(* IEC 61131-3 sources: Aqueous_Solutions/docs-authority/plc (part 2) *)

(* ---- PLC-FAB.st ---- *)
(* AQS-CTL-004 X-CTL-04: control program source, generated by flow_graph/control/plc_programs.py *)
(* Basis: AQS-CTL-001 INSTRUMENT_INDEX.csv, AQS-CTL-002 control architecture, graph set-points. *)
(* PLC-FAB: CPU single; IO counts AI 72 AO 3 DI 92 DO 13 (modules per AQS-CTL-002, 16-channel, 20 % spare) *)
PROGRAM PLC_FAB_CTRL
VAR
  (* 100 ms cyclic task per AQS-CTL-002 *)
  WAFER_FABFT-01_PV : REAL ;  (* S39 normal 0.14 L/h )
  WAFER_FABFT-02_PV : REAL ;  (* S39B normal 0.00 L/h )
  WAFER_FABFT-03_PV : REAL ;  (* IA-FAB-SPENT normal 2.77 L/h )
  WAFER_FABFT-04_PV : REAL ;  (* IA-FAB-N2-VENT normal 0.03 L/h )
  WAFER_FABFT-05_PV : REAL ;  (* IA-AR-CZ-BACK normal 0.14 L/h )
  WAFER_FABLT-01_PV : REAL ;  (* A-M-182 liquid height )
  WAFER_FABPT-01_PV : REAL ;  (* no design pressure on the graph )
  WAFER_FABTE-01_PV : REAL ;  (* band by service )
  WET_BENCHFT-01_PV : REAL ;  (* S10 normal 3.29 L/h )
  WET_BENCHFT-02_PV : REAL ;  (* S38 normal 0.00 L/h )
  WET_BENCHLT-01_PV : REAL ;  (* A-M-182 liquid height )
  WET_BENCHPT-01_PV : REAL ;  (* no design pressure on the graph )
  WET_BENCHTE-01_PV : REAL ;  (* band by service )
  LITHO_ALIGNPT-01_PV : REAL ;  (* no design pressure on the graph )
  LITHO_ALIGNTE-01_PV : REAL ;  (* band by service )
  LITHO_COATPT-01_PV : REAL ;  (* no design pressure on the graph )
  LITHO_COATTE-01_PV : REAL ;  (* band by service )
  RESIST_SYNLT-01_PV : REAL ;  (* A-M-182 liquid height )
  RESIST_SYNPT-01_PV : REAL ;  (* no design pressure on the graph )
  RESIST_SYNTE-01_PV : REAL ;  (* band by service )
  SOLV_PLANTLT-01_PV : REAL ;  (* A-M-182 liquid height )
  SOLV_PLANTPT-01_PV : REAL ;  (* no design pressure on the graph )
  SOLV_PLANTTE-01_PV : REAL ;  (* band by service )
  WS_AMMONIAFT-01_PV : REAL ;  (* S33 normal 0.13 L/h )
  WS_AMMONIAFT-02_PV : REAL ;  (* IA-NH3-MET normal 0.00 L/h )
  WS_AMMONIALT-01_PV : REAL ;  (* A-M-182 liquid height )
  WS_AMMONIAPT-01_PV : REAL ;  (* no design pressure on the graph )
  WS_AMMONIATE-01_PV : REAL ;  (* band by service )
  WS_DOPELT-01_PV : REAL ;  (* A-M-182 liquid height )
  WS_DOPEPT-01_PV : REAL ;  (* no design pressure on the graph )
  WS_DOPETE-01_PV : REAL ;  (* band by service )
  WS_HF_EDFT-01_PV : REAL ;  (* S31 normal 0.06 L/h )
  WS_HF_EDLT-01_PV : REAL ;  (* A-M-182 liquid height )
  WS_HF_EDPT-01_PV : REAL ;  (* no design pressure on the graph )
  WS_HF_EDTE-01_PV : REAL ;  (* band by service )
  WS_KOHFT-01_PV : REAL ;  (* S35 normal 0.01 L/h )
  WS_KOHLT-01_PV : REAL ;  (* A-M-182 liquid height )
  WS_KOHPT-01_PV : REAL ;  (* no design pressure on the graph )
  WS_KOHTE-01_PV : REAL ;  (* band by service )
  WS_NITRICFT-01_PV : REAL ;  (* S34 normal 0.05 L/h )
  WS_NITRICFT-02_PV : REAL ;  (* IA-NIT-VENT normal 0.00 L/h )
  WS_NITRICLT-01_PV : REAL ;  (* A-M-182 liquid height )
  WS_NITRICPT-01_PV : REAL ;  (* no design pressure on the graph )
  WS_NITRICTE-01_PV : REAL ;  (* band by service )
  WS_PEROXFT-01_PV : REAL ;  (* S32 normal 0.12 L/h )
  WS_PEROXLT-01_PV : REAL ;  (* A-M-182 liquid height )
  WS_PEROXPT-01_PV : REAL ;  (* no design pressure on the graph )
  WS_PEROXTE-01_PV : REAL ;  (* band by service )
  WS_PHOSFT-01_PV : REAL ;  (* S34B normal 0.03 L/h )
  WS_PHOSFT-02_PV : REAL ;  (* IA-PHOS-DOPE normal 0.00 L/h )
  WS_PHOSLT-01_PV : REAL ;  (* A-M-182 liquid height )
  WS_PHOSPT-01_PV : REAL ;  (* no design pressure on the graph )
  WS_PHOSTE-01_PV : REAL ;  (* band by service )
  WS_SLURRYFT-01_PV : REAL ;  (* S37 normal 0.14 L/h )
  WS_SLURRYLT-01_PV : REAL ;  (* A-M-182 liquid height )
  WS_SLURRYPT-01_PV : REAL ;  (* no design pressure on the graph )
  WS_SLURRYTE-01_PV : REAL ;  (* band by service )
  WS_SOLVFT-01_PV : REAL ;  (* IA-SOLV-WB normal 0.01 L/h )
  WS_SOLVFT-02_PV : REAL ;  (* IA-FAB-SOLV normal 0.00 L/h )
  WS_SOLVLT-01_PV : REAL ;  (* A-M-182 liquid height )
  WS_SOLVPT-01_PV : REAL ;  (* no design pressure on the graph )
  WS_SOLVTE-01_PV : REAL ;  (* band by service )
  LITHO_STUBPT-01_PV : REAL ;  (* no design pressure on the graph )
  LITHO_STUBTE-01_PV : REAL ;  (* band by service )
  FAB_UPW_TANKFT-01_PV : REAL ;  (* S27 normal 2.50 L/h )
  FAB_UPW_TANKLT-01_PV : REAL ;  (* A-M-182 liquid height )
  FAB_UPW_TANKPT-01_PV : REAL ;  (* no design pressure on the graph )
  FAB_UPW_TANKTE-01_PV : REAL ;  (* band by service )
  SOLAR_PV_CELLPT-01_PV : REAL ;  (* no design pressure on the graph )
  SOLAR_PV_CELLTE-01_PV : REAL ;  (* band by service )
  LITHO_DEVPT-01_PV : REAL ;  (* no design pressure on the graph )
  LITHO_DEVTE-01_PV : REAL ;  (* band by service )
END_VAR

  (* FLOW control loop - set-point from the graph basis *)
  WAFER_FABFT-01_SP := 0.14 ;  (* graph basis: S39 normal 0.14 L/h )
  FB_PI_WAFER_FABFT-01( PV := WAFER_FABFT-01_PV, SP := WAFER_FABFT-01_SP );  (* PI per AQS-CTL-002; GAIN/KI entered at commissioning from the step test (AQS-COM-001 sec. 3), anti-windup clamp per this FB *)
  WAFER_FABFT-01_ALARM_HI := 0.15400000000000003 ;  (* SP x 1.1 margin, A-M-188 margin class *)
  WAFER_FABFT-01_ALARM_LO := 0.12600000000000003 ;

  (* FLOW control loop - set-point from the graph basis *)
  WAFER_FABFT-02_SP := 0.0 ;  (* graph basis: S39B normal 0.00 L/h )
  FB_PI_WAFER_FABFT-02( PV := WAFER_FABFT-02_PV, SP := WAFER_FABFT-02_SP );  (* PI per AQS-CTL-002; GAIN/KI entered at commissioning from the step test (AQS-COM-001 sec. 3), anti-windup clamp per this FB *)
  WAFER_FABFT-02_ALARM_HI := 0.0 ;  (* expected-zero state: any positive PV alarms )

  (* FLOW control loop - set-point from the graph basis *)
  WAFER_FABFT-03_SP := 2.77 ;  (* graph basis: IA-FAB-SPENT normal 2.77 L/h )
  FB_PI_WAFER_FABFT-03( PV := WAFER_FABFT-03_PV, SP := WAFER_FABFT-03_SP );  (* PI per AQS-CTL-002; GAIN/KI entered at commissioning from the step test (AQS-COM-001 sec. 3), anti-windup clamp per this FB *)
  WAFER_FABFT-03_ALARM_HI := 3.047 ;  (* SP x 1.1 margin, A-M-188 margin class *)
  WAFER_FABFT-03_ALARM_LO := 2.493 ;

  (* FLOW control loop - set-point from the graph basis *)
  WAFER_FABFT-04_SP := 0.03 ;  (* graph basis: IA-FAB-N2-VENT normal 0.03 L/h )
  FB_PI_WAFER_FABFT-04( PV := WAFER_FABFT-04_PV, SP := WAFER_FABFT-04_SP );  (* PI per AQS-CTL-002; GAIN/KI entered at commissioning from the step test (AQS-COM-001 sec. 3), anti-windup clamp per this FB *)
  WAFER_FABFT-04_ALARM_HI := 0.033 ;  (* SP x 1.1 margin, A-M-188 margin class *)
  WAFER_FABFT-04_ALARM_LO := 0.027 ;

  (* FLOW control loop - set-point from the graph basis *)
  WAFER_FABFT-05_SP := 0.14 ;  (* graph basis: IA-AR-CZ-BACK normal 0.14 L/h )
  FB_PI_WAFER_FABFT-05( PV := WAFER_FABFT-05_PV, SP := WAFER_FABFT-05_SP );  (* PI per AQS-CTL-002; GAIN/KI entered at commissioning from the step test (AQS-COM-001 sec. 3), anti-windup clamp per this FB *)
  WAFER_FABFT-05_ALARM_HI := 0.15400000000000003 ;  (* SP x 1.1 margin, A-M-188 margin class *)
  WAFER_FABFT-05_ALARM_LO := 0.12600000000000003 ;

  (* LEVEL monitoring block - indication, no set-point invented )
  FB_AI_WAFER_FABLT-01( PV := WAFER_FABLT-01_PV );
  WAFER_FABLT-01_ALARM_HI := 90.0 ;  (* 90 % of span, registered LSH convention )

  (* PRESSURE monitoring block - indication, no set-point invented )
  FB_AI_WAFER_FABPT-01( PV := WAFER_FABPT-01_PV );
  WAFER_FABPT-01_ALARM_HI := 9.0 ;  (* 90 % of span, registered LSH convention )

  (* TEMPERATURE monitoring block - indication, no set-point invented )
  FB_AI_WAFER_FABTE-01( PV := WAFER_FABTE-01_PV );
  WAFER_FABTE-01_ALARM_HI := 135.0 ;  (* 90 % of span, registered LSH convention )

  (* FLOW control loop - set-point from the graph basis *)
  WET_BENCHFT-01_SP := 3.29 ;  (* graph basis: S10 normal 3.29 L/h )
  FB_PI_WET_BENCHFT-01( PV := WET_BENCHFT-01_PV, SP := WET_BENCHFT-01_SP );  (* PI per AQS-CTL-002; GAIN/KI entered at commissioning from the step test (AQS-COM-001 sec. 3), anti-windup clamp per this FB *)
  WET_BENCHFT-01_ALARM_HI := 3.619 ;  (* SP x 1.1 margin, A-M-188 margin class *)
  WET_BENCHFT-01_ALARM_LO := 2.9610000000000003 ;

  (* FLOW control loop - set-point from the graph basis *)
  WET_BENCHFT-02_SP := 0.0 ;  (* graph basis: S38 normal 0.00 L/h )
  FB_PI_WET_BENCHFT-02( PV := WET_BENCHFT-02_PV, SP := WET_BENCHFT-02_SP );  (* PI per AQS-CTL-002; GAIN/KI entered at commissioning from the step test (AQS-COM-001 sec. 3), anti-windup clamp per this FB *)
  WET_BENCHFT-02_ALARM_HI := 0.0 ;  (* expected-zero state: any positive PV alarms )

  (* LEVEL monitoring block - indication, no set-point invented )
  FB_AI_WET_BENCHLT-01( PV := WET_BENCHLT-01_PV );
  WET_BENCHLT-01_ALARM_HI := 90.0 ;  (* 90 % of span, registered LSH convention )

  (* PRESSURE monitoring block - indication, no set-point invented )
  FB_AI_WET_BENCHPT-01( PV := WET_BENCHPT-01_PV );
  WET_BENCHPT-01_ALARM_HI := 9.0 ;  (* 90 % of span, registered LSH convention )

  (* TEMPERATURE monitoring block - indication, no set-point invented )
  FB_AI_WET_BENCHTE-01( PV := WET_BENCHTE-01_PV );
  WET_BENCHTE-01_ALARM_HI := 135.0 ;  (* 90 % of span, registered LSH convention )

  (* PRESSURE monitoring block - indication, no set-point invented )
  FB_AI_LITHO_ALIGNPT-01( PV := LITHO_ALIGNPT-01_PV );
  LITHO_ALIGNPT-01_ALARM_HI := 9.0 ;  (* 90 % of span, registered LSH convention )

  (* TEMPERATURE monitoring block - indication, no set-point invented )
  FB_AI_LITHO_ALIGNTE-01( PV := LITHO_ALIGNTE-01_PV );
  LITHO_ALIGNTE-01_ALARM_HI := 135.0 ;  (* 90 % of span, registered LSH convention )

  (* PRESSURE monitoring block - indication, no set-point invented )
  FB_AI_LITHO_COATPT-01( PV := LITHO_COATPT-01_PV );
  LITHO_COATPT-01_ALARM_HI := 9.0 ;  (* 90 % of span, registered LSH convention )

  (* TEMPERATURE monitoring block - indication, no set-point invented )
  FB_AI_LITHO_COATTE-01( PV := LITHO_COATTE-01_PV );
  LITHO_COATTE-01_ALARM_HI := 135.0 ;  (* 90 % of span, registered LSH convention )

  (* LEVEL monitoring block - indication, no set-point invented )
  FB_AI_RESIST_SYNLT-01( PV := RESIST_SYNLT-01_PV );
  RESIST_SYNLT-01_ALARM_HI := 90.0 ;  (* 90 % of span, registered LSH convention )

  (* PRESSURE monitoring block - indication, no set-point invented )
  FB_AI_RESIST_SYNPT-01( PV := RESIST_SYNPT-01_PV );
  RESIST_SYNPT-01_ALARM_HI := 9.0 ;  (* 90 % of span, registered LSH convention )

  (* TEMPERATURE monitoring block - indication, no set-point invented )
  FB_AI_RESIST_SYNTE-01( PV := RESIST_SYNTE-01_PV );
  RESIST_SYNTE-01_ALARM_HI := 135.0 ;  (* 90 % of span, registered LSH convention )

  (* LEVEL monitoring block - indication, no set-point invented )
  FB_AI_SOLV_PLANTLT-01( PV := SOLV_PLANTLT-01_PV );
  SOLV_PLANTLT-01_ALARM_HI := 90.0 ;  (* 90 % of span, registered LSH convention )

  (* PRESSURE monitoring block - indication, no set-point invented )
  FB_AI_SOLV_PLANTPT-01( PV := SOLV_PLANTPT-01_PV );
  SOLV_PLANTPT-01_ALARM_HI := 9.0 ;  (* 90 % of span, registered LSH convention )

  (* TEMPERATURE monitoring block - indication, no set-point invented )
  FB_AI_SOLV_PLANTTE-01( PV := SOLV_PLANTTE-01_PV );
  SOLV_PLANTTE-01_ALARM_HI := 135.0 ;  (* 90 % of span, registered LSH convention )

  (* FLOW control loop - set-point from the graph basis *)
  WS_AMMONIAFT-01_SP := 0.13 ;  (* graph basis: S33 normal 0.13 L/h )
  FB_PI_WS_AMMONIAFT-01( PV := WS_AMMONIAFT-01_PV, SP := WS_AMMONIAFT-01_SP );  (* PI per AQS-CTL-002; GAIN/KI entered at commissioning from the step test (AQS-COM-001 sec. 3), anti-windup clamp per this FB *)
  WS_AMMONIAFT-01_ALARM_HI := 0.14300000000000002 ;  (* SP x 1.1 margin, A-M-188 margin class *)
  WS_AMMONIAFT-01_ALARM_LO := 0.117 ;

  (* FLOW control loop - set-point from the graph basis *)
  WS_AMMONIAFT-02_SP := 0.0 ;  (* graph basis: IA-NH3-MET normal 0.00 L/h )
  FB_PI_WS_AMMONIAFT-02( PV := WS_AMMONIAFT-02_PV, SP := WS_AMMONIAFT-02_SP );  (* PI per AQS-CTL-002; GAIN/KI entered at commissioning from the step test (AQS-COM-001 sec. 3), anti-windup clamp per this FB *)
  WS_AMMONIAFT-02_ALARM_HI := 0.0 ;  (* expected-zero state: any positive PV alarms )

  (* LEVEL monitoring block - indication, no set-point invented )
  FB_AI_WS_AMMONIALT-01( PV := WS_AMMONIALT-01_PV );
  WS_AMMONIALT-01_ALARM_HI := 90.0 ;  (* 90 % of span, registered LSH convention )

  (* PRESSURE monitoring block - indication, no set-point invented )
  FB_AI_WS_AMMONIAPT-01( PV := WS_AMMONIAPT-01_PV );
  WS_AMMONIAPT-01_ALARM_HI := 9.0 ;  (* 90 % of span, registered LSH convention )

  (* TEMPERATURE monitoring block - indication, no set-point invented )
  FB_AI_WS_AMMONIATE-01( PV := WS_AMMONIATE-01_PV );
  WS_AMMONIATE-01_ALARM_HI := 135.0 ;  (* 90 % of span, registered LSH convention )

  (* LEVEL monitoring block - indication, no set-point invented )
  FB_AI_WS_DOPELT-01( PV := WS_DOPELT-01_PV );
  WS_DOPELT-01_ALARM_HI := 90.0 ;  (* 90 % of span, registered LSH convention )

  (* PRESSURE monitoring block - indication, no set-point invented )
  FB_AI_WS_DOPEPT-01( PV := WS_DOPEPT-01_PV );
  WS_DOPEPT-01_ALARM_HI := 9.0 ;  (* 90 % of span, registered LSH convention )

  (* TEMPERATURE monitoring block - indication, no set-point invented )
  FB_AI_WS_DOPETE-01( PV := WS_DOPETE-01_PV );
  WS_DOPETE-01_ALARM_HI := 135.0 ;  (* 90 % of span, registered LSH convention )

  (* FLOW control loop - set-point from the graph basis *)
  WS_HF_EDFT-01_SP := 0.06 ;  (* graph basis: S31 normal 0.06 L/h )
  FB_PI_WS_HF_EDFT-01( PV := WS_HF_EDFT-01_PV, SP := WS_HF_EDFT-01_SP );  (* PI per AQS-CTL-002; GAIN/KI entered at commissioning from the step test (AQS-COM-001 sec. 3), anti-windup clamp per this FB *)
  WS_HF_EDFT-01_ALARM_HI := 0.066 ;  (* SP x 1.1 margin, A-M-188 margin class *)
  WS_HF_EDFT-01_ALARM_LO := 0.054 ;

  (* LEVEL monitoring block - indication, no set-point invented )
  FB_AI_WS_HF_EDLT-01( PV := WS_HF_EDLT-01_PV );
  WS_HF_EDLT-01_ALARM_HI := 90.0 ;  (* 90 % of span, registered LSH convention )

  (* PRESSURE monitoring block - indication, no set-point invented )
  FB_AI_WS_HF_EDPT-01( PV := WS_HF_EDPT-01_PV );
  WS_HF_EDPT-01_ALARM_HI := 9.0 ;  (* 90 % of span, registered LSH convention )

  (* TEMPERATURE monitoring block - indication, no set-point invented )
  FB_AI_WS_HF_EDTE-01( PV := WS_HF_EDTE-01_PV );
  WS_HF_EDTE-01_ALARM_HI := 135.0 ;  (* 90 % of span, registered LSH convention )

  (* FLOW control loop - set-point from the graph basis *)
  WS_KOHFT-01_SP := 0.01 ;  (* graph basis: S35 normal 0.01 L/h )
  FB_PI_WS_KOHFT-01( PV := WS_KOHFT-01_PV, SP := WS_KOHFT-01_SP );  (* PI per AQS-CTL-002; GAIN/KI entered at commissioning from the step test (AQS-COM-001 sec. 3), anti-windup clamp per this FB *)
  WS_KOHFT-01_ALARM_HI := 0.011000000000000001 ;  (* SP x 1.1 margin, A-M-188 margin class *)
  WS_KOHFT-01_ALARM_LO := 0.009000000000000001 ;

  (* LEVEL monitoring block - indication, no set-point invented )
  FB_AI_WS_KOHLT-01( PV := WS_KOHLT-01_PV );
  WS_KOHLT-01_ALARM_HI := 90.0 ;  (* 90 % of span, registered LSH convention )

  (* PRESSURE monitoring block - indication, no set-point invented )
  FB_AI_WS_KOHPT-01( PV := WS_KOHPT-01_PV );
  WS_KOHPT-01_ALARM_HI := 9.0 ;  (* 90 % of span, registered LSH convention )

  (* TEMPERATURE monitoring block - indication, no set-point invented )
  FB_AI_WS_KOHTE-01( PV := WS_KOHTE-01_PV );
  WS_KOHTE-01_ALARM_HI := 135.0 ;  (* 90 % of span, registered LSH convention )

  (* FLOW control loop - set-point from the graph basis *)
  WS_NITRICFT-01_SP := 0.05 ;  (* graph basis: S34 normal 0.05 L/h )
  FB_PI_WS_NITRICFT-01( PV := WS_NITRICFT-01_PV, SP := WS_NITRICFT-01_SP );  (* PI per AQS-CTL-002; GAIN/KI entered at commissioning from the step test (AQS-COM-001 sec. 3), anti-windup clamp per this FB *)
  WS_NITRICFT-01_ALARM_HI := 0.05500000000000001 ;  (* SP x 1.1 margin, A-M-188 margin class *)
  WS_NITRICFT-01_ALARM_LO := 0.045000000000000005 ;

  (* FLOW control loop - set-point from the graph basis *)
  WS_NITRICFT-02_SP := 0.0 ;  (* graph basis: IA-NIT-VENT normal 0.00 L/h )
  FB_PI_WS_NITRICFT-02( PV := WS_NITRICFT-02_PV, SP := WS_NITRICFT-02_SP );  (* PI per AQS-CTL-002; GAIN/KI entered at commissioning from the step test (AQS-COM-001 sec. 3), anti-windup clamp per this FB *)
  WS_NITRICFT-02_ALARM_HI := 0.0 ;  (* expected-zero state: any positive PV alarms )

  (* LEVEL monitoring block - indication, no set-point invented )
  FB_AI_WS_NITRICLT-01( PV := WS_NITRICLT-01_PV );
  WS_NITRICLT-01_ALARM_HI := 90.0 ;  (* 90 % of span, registered LSH convention )

  (* PRESSURE monitoring block - indication, no set-point invented )
  FB_AI_WS_NITRICPT-01( PV := WS_NITRICPT-01_PV );
  WS_NITRICPT-01_ALARM_HI := 9.0 ;  (* 90 % of span, registered LSH convention )

  (* TEMPERATURE monitoring block - indication, no set-point invented )
  FB_AI_WS_NITRICTE-01( PV := WS_NITRICTE-01_PV );
  WS_NITRICTE-01_ALARM_HI := 135.0 ;  (* 90 % of span, registered LSH convention )

  (* FLOW control loop - set-point from the graph basis *)
  WS_PEROXFT-01_SP := 0.12 ;  (* graph basis: S32 normal 0.12 L/h )
  FB_PI_WS_PEROXFT-01( PV := WS_PEROXFT-01_PV, SP := WS_PEROXFT-01_SP );  (* PI per AQS-CTL-002; GAIN/KI entered at commissioning from the step test (AQS-COM-001 sec. 3), anti-windup clamp per this FB *)
  WS_PEROXFT-01_ALARM_HI := 0.132 ;  (* SP x 1.1 margin, A-M-188 margin class *)
  WS_PEROXFT-01_ALARM_LO := 0.108 ;

  (* LEVEL monitoring block - indication, no set-point invented )
  FB_AI_WS_PEROXLT-01( PV := WS_PEROXLT-01_PV );
  WS_PEROXLT-01_ALARM_HI := 90.0 ;  (* 90 % of span, registered LSH convention )

  (* PRESSURE monitoring block - indication, no set-point invented )
  FB_AI_WS_PEROXPT-01( PV := WS_PEROXPT-01_PV );
  WS_PEROXPT-01_ALARM_HI := 9.0 ;  (* 90 % of span, registered LSH convention )

  (* TEMPERATURE monitoring block - indication, no set-point invented )
  FB_AI_WS_PEROXTE-01( PV := WS_PEROXTE-01_PV );
  WS_PEROXTE-01_ALARM_HI := 135.0 ;  (* 90 % of span, registered LSH convention )

  (* FLOW control loop - set-point from the graph basis *)
  WS_PHOSFT-01_SP := 0.03 ;  (* graph basis: S34B normal 0.03 L/h )
  FB_PI_WS_PHOSFT-01( PV := WS_PHOSFT-01_PV, SP := WS_PHOSFT-01_SP );  (* PI per AQS-CTL-002; GAIN/KI entered at commissioning from the step test (AQS-COM-001 sec. 3), anti-windup clamp per this FB *)
  WS_PHOSFT-01_ALARM_HI := 0.033 ;  (* SP x 1.1 margin, A-M-188 margin class *)
  WS_PHOSFT-01_ALARM_LO := 0.027 ;

  (* FLOW control loop - set-point from the graph basis *)
  WS_PHOSFT-02_SP := 0.0 ;  (* graph basis: IA-PHOS-DOPE normal 0.00 L/h )
  FB_PI_WS_PHOSFT-02( PV := WS_PHOSFT-02_PV, SP := WS_PHOSFT-02_SP );  (* PI per AQS-CTL-002; GAIN/KI entered at commissioning from the step test (AQS-COM-001 sec. 3), anti-windup clamp per this FB *)
  WS_PHOSFT-02_ALARM_HI := 0.0 ;  (* expected-zero state: any positive PV alarms )

  (* LEVEL monitoring block - indication, no set-point invented )
  FB_AI_WS_PHOSLT-01( PV := WS_PHOSLT-01_PV );
  WS_PHOSLT-01_ALARM_HI := 90.0 ;  (* 90 % of span, registered LSH convention )

  (* PRESSURE monitoring block - indication, no set-point invented )
  FB_AI_WS_PHOSPT-01( PV := WS_PHOSPT-01_PV );
  WS_PHOSPT-01_ALARM_HI := 9.0 ;  (* 90 % of span, registered LSH convention )

  (* TEMPERATURE monitoring block - indication, no set-point invented )
  FB_AI_WS_PHOSTE-01( PV := WS_PHOSTE-01_PV );
  WS_PHOSTE-01_ALARM_HI := 135.0 ;  (* 90 % of span, registered LSH convention )

  (* FLOW control loop - set-point from the graph basis *)
  WS_SLURRYFT-01_SP := 0.14 ;  (* graph basis: S37 normal 0.14 L/h )
  FB_PI_WS_SLURRYFT-01( PV := WS_SLURRYFT-01_PV, SP := WS_SLURRYFT-01_SP );  (* PI per AQS-CTL-002; GAIN/KI entered at commissioning from the step test (AQS-COM-001 sec. 3), anti-windup clamp per this FB *)
  WS_SLURRYFT-01_ALARM_HI := 0.15400000000000003 ;  (* SP x 1.1 margin, A-M-188 margin class *)
  WS_SLURRYFT-01_ALARM_LO := 0.12600000000000003 ;

  (* LEVEL monitoring block - indication, no set-point invented )
  FB_AI_WS_SLURRYLT-01( PV := WS_SLURRYLT-01_PV );
  WS_SLURRYLT-01_ALARM_HI := 90.0 ;  (* 90 % of span, registered LSH convention )

  (* PRESSURE monitoring block - indication, no set-point invented )
  FB_AI_WS_SLURRYPT-01( PV := WS_SLURRYPT-01_PV );
  WS_SLURRYPT-01_ALARM_HI := 9.0 ;  (* 90 % of span, registered LSH convention )

  (* TEMPERATURE monitoring block - indication, no set-point invented )
  FB_AI_WS_SLURRYTE-01( PV := WS_SLURRYTE-01_PV );
  WS_SLURRYTE-01_ALARM_HI := 135.0 ;  (* 90 % of span, registered LSH convention )

  (* FLOW control loop - set-point from the graph basis *)
  WS_SOLVFT-01_SP := 0.01 ;  (* graph basis: IA-SOLV-WB normal 0.01 L/h )
  FB_PI_WS_SOLVFT-01( PV := WS_SOLVFT-01_PV, SP := WS_SOLVFT-01_SP );  (* PI per AQS-CTL-002; GAIN/KI entered at commissioning from the step test (AQS-COM-001 sec. 3), anti-windup clamp per this FB *)
  WS_SOLVFT-01_ALARM_HI := 0.011000000000000001 ;  (* SP x 1.1 margin, A-M-188 margin class *)
  WS_SOLVFT-01_ALARM_LO := 0.009000000000000001 ;

  (* FLOW control loop - set-point from the graph basis *)
  WS_SOLVFT-02_SP := 0.0 ;  (* graph basis: IA-FAB-SOLV normal 0.00 L/h )
  FB_PI_WS_SOLVFT-02( PV := WS_SOLVFT-02_PV, SP := WS_SOLVFT-02_SP );  (* PI per AQS-CTL-002; GAIN/KI entered at commissioning from the step test (AQS-COM-001 sec. 3), anti-windup clamp per this FB *)
  WS_SOLVFT-02_ALARM_HI := 0.0 ;  (* expected-zero state: any positive PV alarms )

  (* LEVEL monitoring block - indication, no set-point invented )
  FB_AI_WS_SOLVLT-01( PV := WS_SOLVLT-01_PV );
  WS_SOLVLT-01_ALARM_HI := 90.0 ;  (* 90 % of span, registered LSH convention )

  (* PRESSURE monitoring block - indication, no set-point invented )
  FB_AI_WS_SOLVPT-01( PV := WS_SOLVPT-01_PV );
  WS_SOLVPT-01_ALARM_HI := 9.0 ;  (* 90 % of span, registered LSH convention )

  (* TEMPERATURE monitoring block - indication, no set-point invented )
  FB_AI_WS_SOLVTE-01( PV := WS_SOLVTE-01_PV );
  WS_SOLVTE-01_ALARM_HI := 135.0 ;  (* 90 % of span, registered LSH convention )

  (* PRESSURE monitoring block - indication, no set-point invented )
  FB_AI_LITHO_STUBPT-01( PV := LITHO_STUBPT-01_PV );
  LITHO_STUBPT-01_ALARM_HI := 9.0 ;  (* 90 % of span, registered LSH convention )

  (* TEMPERATURE monitoring block - indication, no set-point invented )
  FB_AI_LITHO_STUBTE-01( PV := LITHO_STUBTE-01_PV );
  LITHO_STUBTE-01_ALARM_HI := 135.0 ;  (* 90 % of span, registered LSH convention )

  (* FLOW control loop - set-point from the graph basis *)
  FAB_UPW_TANKFT-01_SP := 2.5 ;  (* graph basis: S27 normal 2.50 L/h )
  FB_PI_FAB_UPW_TANKFT-01( PV := FAB_UPW_TANKFT-01_PV, SP := FAB_UPW_TANKFT-01_SP );  (* PI per AQS-CTL-002; GAIN/KI entered at commissioning from the step test (AQS-COM-001 sec. 3), anti-windup clamp per this FB *)
  FAB_UPW_TANKFT-01_ALARM_HI := 2.75 ;  (* SP x 1.1 margin, A-M-188 margin class *)
  FAB_UPW_TANKFT-01_ALARM_LO := 2.25 ;

  (* LEVEL monitoring block - indication, no set-point invented )
  FB_AI_FAB_UPW_TANKLT-01( PV := FAB_UPW_TANKLT-01_PV );
  FAB_UPW_TANKLT-01_ALARM_HI := 90.0 ;  (* 90 % of span, registered LSH convention )

  (* PRESSURE monitoring block - indication, no set-point invented )
  FB_AI_FAB_UPW_TANKPT-01( PV := FAB_UPW_TANKPT-01_PV );
  FAB_UPW_TANKPT-01_ALARM_HI := 9.0 ;  (* 90 % of span, registered LSH convention )

  (* TEMPERATURE monitoring block - indication, no set-point invented )
  FB_AI_FAB_UPW_TANKTE-01( PV := FAB_UPW_TANKTE-01_PV );
  FAB_UPW_TANKTE-01_ALARM_HI := 135.0 ;  (* 90 % of span, registered LSH convention )

  (* PRESSURE monitoring block - indication, no set-point invented )
  FB_AI_SOLAR_PV_CELLPT-01( PV := SOLAR_PV_CELLPT-01_PV );
  SOLAR_PV_CELLPT-01_ALARM_HI := 9.0 ;  (* 90 % of span, registered LSH convention )

  (* TEMPERATURE monitoring block - indication, no set-point invented )
  FB_AI_SOLAR_PV_CELLTE-01( PV := SOLAR_PV_CELLTE-01_PV );
  SOLAR_PV_CELLTE-01_ALARM_HI := 135.0 ;  (* 90 % of span, registered LSH convention )

  (* PRESSURE monitoring block - indication, no set-point invented )
  FB_AI_LITHO_DEVPT-01( PV := LITHO_DEVPT-01_PV );
  LITHO_DEVPT-01_ALARM_HI := 9.0 ;  (* 90 % of span, registered LSH convention )

  (* TEMPERATURE monitoring block - indication, no set-point invented )
  FB_AI_LITHO_DEVTE-01( PV := LITHO_DEVTE-01_PV );
  LITHO_DEVTE-01_ALARM_HI := 135.0 ;  (* 90 % of span, registered LSH convention )

END_PROGRAM

(* ---- PLC-FARM.st ---- *)
(* AQS-CTL-004 X-CTL-04: control program source, generated by flow_graph/control/plc_programs.py *)
(* Basis: AQS-CTL-001 INSTRUMENT_INDEX.csv, AQS-CTL-002 control architecture, graph set-points. *)
(* PLC-FARM: CPU redundant pair; IO counts AI 48 AO 0 DI 3 DO 0 (modules per AQS-CTL-002, 16-channel, 20 % spare) *)
PROGRAM PLC_FARM_CTRL
VAR
  (* 100 ms cyclic task per AQS-CTL-002 *)
  GROW_BEDFT-01_PV : REAL ;  (* S13 normal 0.16 L/h )
  GROW_BEDFT-02_PV : REAL ;  (* S15 normal 0.00 L/h )
  GROW_BEDFT-03_PV : REAL ;  (* S87 normal 0.03 L/h )
  GROW_BEDFT-04_PV : REAL ;  (* FARM_O2_TO_HAB normal 0.00 L/h )
  GROW_BEDFT-05_PV : REAL ;  (* IA-BED-VAP normal 2.81 L/h )
  GROW_BEDFT-06_PV : REAL ;  (* RABBIT_FORAGE normal 0.02 L/h )
  GROW_BEDFT-07_PV : REAL ;  (* NECTAR_FORAGE normal 0.01 L/h )
  GROW_BEDFT-08_PV : REAL ;  (* VERMI_FEED normal 0.04 L/h )
  GROW_BEDLT-01_PV : REAL ;  (* A-M-182 liquid height )
  GROW_BEDPT-01_PV : REAL ;  (* no design pressure on the graph )
  GROW_BEDTE-01_PV : REAL ;  (* band by service )
  DUCKWEEDPT-01_PV : REAL ;  (* no design pressure on the graph )
  DUCKWEEDTE-01_PV : REAL ;  (* band by service )
  BIOFILTERPT-01_PV : REAL ;  (* no design pressure on the graph )
  BIOFILTERTE-01_PV : REAL ;  (* band by service )
  BSFL_BINPT-01_PV : REAL ;  (* no design pressure on the graph )
  BSFL_BINTE-01_PV : REAL ;  (* band by service )
  QUAIL_CAGEPT-01_PV : REAL ;  (* no design pressure on the graph )
  QUAIL_CAGETE-01_PV : REAL ;  (* band by service )
  CHICKEN_COOPPT-01_PV : REAL ;  (* no design pressure on the graph )
  CHICKEN_COOPTE-01_PV : REAL ;  (* band by service )
  FEED_PREPPT-01_PV : REAL ;  (* no design pressure on the graph )
  FEED_PREPTE-01_PV : REAL ;  (* band by service )
  AQUA_TANKPT-01_PV : REAL ;  (* no design pressure on the graph )
  AQUA_TANKTE-01_PV : REAL ;  (* band by service )
  GROWBED_APT-01_PV : REAL ;  (* no design pressure on the graph )
  GROWBED_ATE-01_PV : REAL ;  (* band by service )
  GROWBED_BPT-01_PV : REAL ;  (* no design pressure on the graph )
  GROWBED_BTE-01_PV : REAL ;  (* band by service )
  BEE_HIVEPT-01_PV : REAL ;  (* no design pressure on the graph )
  BEE_HIVETE-01_PV : REAL ;  (* band by service )
  RABBIT_HUTCHPT-01_PV : REAL ;  (* no design pressure on the graph )
  RABBIT_HUTCHTE-01_PV : REAL ;  (* band by service )
  DUCK_PENPT-01_PV : REAL ;  (* no design pressure on the graph )
  DUCK_PENTE-01_PV : REAL ;  (* band by service )
  FOOD_STOREPT-01_PV : REAL ;  (* no design pressure on the graph )
  FOOD_STORETE-01_PV : REAL ;  (* band by service )
  AQUA_UVPT-01_PV : REAL ;  (* no design pressure on the graph )
  AQUA_UVTE-01_PV : REAL ;  (* band by service )
  VERMI_BINPT-01_PV : REAL ;  (* no design pressure on the graph )
  VERMI_BINTE-01_PV : REAL ;  (* band by service )
  FOOD_STORELT-01_PV : REAL ;  (* food stock level: S14 4.2 kg/d )
  HYDRO_GROWAE-01_PV : REAL ;  (* chamber CO2 watch against the habitat management set-point (X-LOC-10 placeholder )
  FEED_PREPPSH-01_PV : REAL ;  (* press-line overpressure interlock on the mash loop (X-FARM-10; A-M-426) )
  AQUA_UVFIT-01_PV : REAL ;  (* loop flow permissive: the UV dose is valid only above the minimum flow (X-FARM-1 )
  AQUA_UVUVT-01_PV : REAL ;  (* dose watchdog: lamp depletion or sleeve fouling decays the signal (X-FARM-12; A- )
  GROWBED_ALT-01_PV : REAL ;  (* flood-and-drain cycle watch on the aerobic root zone (X-FARM build-out; A-M-229) )
  GROWBED_BLT-01_PV : REAL ;  (* mineralisation-zone level watch (X-FARM build-out; A-M-229) )
END_VAR

  (* FLOW control loop - set-point from the graph basis *)
  GROW_BEDFT-01_SP := 0.16 ;  (* graph basis: S13 normal 0.16 L/h )
  FB_PI_GROW_BEDFT-01( PV := GROW_BEDFT-01_PV, SP := GROW_BEDFT-01_SP );  (* PI per AQS-CTL-002; GAIN/KI entered at commissioning from the step test (AQS-COM-001 sec. 3), anti-windup clamp per this FB *)
  GROW_BEDFT-01_ALARM_HI := 0.17600000000000002 ;  (* SP x 1.1 margin, A-M-188 margin class *)
  GROW_BEDFT-01_ALARM_LO := 0.14400000000000002 ;

  (* FLOW control loop - set-point from the graph basis *)
  GROW_BEDFT-02_SP := 0.0 ;  (* graph basis: S15 normal 0.00 L/h )
  FB_PI_GROW_BEDFT-02( PV := GROW_BEDFT-02_PV, SP := GROW_BEDFT-02_SP );  (* PI per AQS-CTL-002; GAIN/KI entered at commissioning from the step test (AQS-COM-001 sec. 3), anti-windup clamp per this FB *)
  GROW_BEDFT-02_ALARM_HI := 0.0 ;  (* expected-zero state: any positive PV alarms )

  (* FLOW control loop - set-point from the graph basis *)
  GROW_BEDFT-03_SP := 0.03 ;  (* graph basis: S87 normal 0.03 L/h )
  FB_PI_GROW_BEDFT-03( PV := GROW_BEDFT-03_PV, SP := GROW_BEDFT-03_SP );  (* PI per AQS-CTL-002; GAIN/KI entered at commissioning from the step test (AQS-COM-001 sec. 3), anti-windup clamp per this FB *)
  GROW_BEDFT-03_ALARM_HI := 0.033 ;  (* SP x 1.1 margin, A-M-188 margin class *)
  GROW_BEDFT-03_ALARM_LO := 0.027 ;

  (* FLOW control loop - set-point from the graph basis *)
  GROW_BEDFT-04_SP := 0.0 ;  (* graph basis: FARM_O2_TO_HAB normal 0.00 L/h )
  FB_PI_GROW_BEDFT-04( PV := GROW_BEDFT-04_PV, SP := GROW_BEDFT-04_SP );  (* PI per AQS-CTL-002; GAIN/KI entered at commissioning from the step test (AQS-COM-001 sec. 3), anti-windup clamp per this FB *)
  GROW_BEDFT-04_ALARM_HI := 0.0 ;  (* expected-zero state: any positive PV alarms )

  (* FLOW control loop - set-point from the graph basis *)
  GROW_BEDFT-05_SP := 2.81 ;  (* graph basis: IA-BED-VAP normal 2.81 L/h )
  FB_PI_GROW_BEDFT-05( PV := GROW_BEDFT-05_PV, SP := GROW_BEDFT-05_SP );  (* PI per AQS-CTL-002; GAIN/KI entered at commissioning from the step test (AQS-COM-001 sec. 3), anti-windup clamp per this FB *)
  GROW_BEDFT-05_ALARM_HI := 3.091 ;  (* SP x 1.1 margin, A-M-188 margin class *)
  GROW_BEDFT-05_ALARM_LO := 2.529 ;

  (* FLOW control loop - set-point from the graph basis *)
  GROW_BEDFT-06_SP := 0.02 ;  (* graph basis: RABBIT_FORAGE normal 0.02 L/h )
  FB_PI_GROW_BEDFT-06( PV := GROW_BEDFT-06_PV, SP := GROW_BEDFT-06_SP );  (* PI per AQS-CTL-002; GAIN/KI entered at commissioning from the step test (AQS-COM-001 sec. 3), anti-windup clamp per this FB *)
  GROW_BEDFT-06_ALARM_HI := 0.022000000000000002 ;  (* SP x 1.1 margin, A-M-188 margin class *)
  GROW_BEDFT-06_ALARM_LO := 0.018000000000000002 ;

  (* FLOW control loop - set-point from the graph basis *)
  GROW_BEDFT-07_SP := 0.01 ;  (* graph basis: NECTAR_FORAGE normal 0.01 L/h )
  FB_PI_GROW_BEDFT-07( PV := GROW_BEDFT-07_PV, SP := GROW_BEDFT-07_SP );  (* PI per AQS-CTL-002; GAIN/KI entered at commissioning from the step test (AQS-COM-001 sec. 3), anti-windup clamp per this FB *)
  GROW_BEDFT-07_ALARM_HI := 0.011000000000000001 ;  (* SP x 1.1 margin, A-M-188 margin class *)
  GROW_BEDFT-07_ALARM_LO := 0.009000000000000001 ;

  (* FLOW control loop - set-point from the graph basis *)
  GROW_BEDFT-08_SP := 0.04 ;  (* graph basis: VERMI_FEED normal 0.04 L/h )
  FB_PI_GROW_BEDFT-08( PV := GROW_BEDFT-08_PV, SP := GROW_BEDFT-08_SP );  (* PI per AQS-CTL-002; GAIN/KI entered at commissioning from the step test (AQS-COM-001 sec. 3), anti-windup clamp per this FB *)
  GROW_BEDFT-08_ALARM_HI := 0.044000000000000004 ;  (* SP x 1.1 margin, A-M-188 margin class *)
  GROW_BEDFT-08_ALARM_LO := 0.036000000000000004 ;

  (* LEVEL monitoring block - indication, no set-point invented )
  FB_AI_GROW_BEDLT-01( PV := GROW_BEDLT-01_PV );
  GROW_BEDLT-01_ALARM_HI := 90.0 ;  (* 90 % of span, registered LSH convention )

  (* PRESSURE monitoring block - indication, no set-point invented )
  FB_AI_GROW_BEDPT-01( PV := GROW_BEDPT-01_PV );
  GROW_BEDPT-01_ALARM_HI := 9.0 ;  (* 90 % of span, registered LSH convention )

  (* TEMPERATURE monitoring block - indication, no set-point invented )
  FB_AI_GROW_BEDTE-01( PV := GROW_BEDTE-01_PV );
  GROW_BEDTE-01_ALARM_HI := 135.0 ;  (* 90 % of span, registered LSH convention )

  (* PRESSURE monitoring block - indication, no set-point invented )
  FB_AI_DUCKWEEDPT-01( PV := DUCKWEEDPT-01_PV );
  DUCKWEEDPT-01_ALARM_HI := 9.0 ;  (* 90 % of span, registered LSH convention )

  (* TEMPERATURE monitoring block - indication, no set-point invented )
  FB_AI_DUCKWEEDTE-01( PV := DUCKWEEDTE-01_PV );
  DUCKWEEDTE-01_ALARM_HI := 135.0 ;  (* 90 % of span, registered LSH convention )

  (* PRESSURE monitoring block - indication, no set-point invented )
  FB_AI_BIOFILTERPT-01( PV := BIOFILTERPT-01_PV );
  BIOFILTERPT-01_ALARM_HI := 9.0 ;  (* 90 % of span, registered LSH convention )

  (* TEMPERATURE monitoring block - indication, no set-point invented )
  FB_AI_BIOFILTERTE-01( PV := BIOFILTERTE-01_PV );
  BIOFILTERTE-01_ALARM_HI := 135.0 ;  (* 90 % of span, registered LSH convention )

  (* PRESSURE monitoring block - indication, no set-point invented )
  FB_AI_BSFL_BINPT-01( PV := BSFL_BINPT-01_PV );
  BSFL_BINPT-01_ALARM_HI := 9.0 ;  (* 90 % of span, registered LSH convention )

  (* TEMPERATURE monitoring block - indication, no set-point invented )
  FB_AI_BSFL_BINTE-01( PV := BSFL_BINTE-01_PV );
  BSFL_BINTE-01_ALARM_HI := 135.0 ;  (* 90 % of span, registered LSH convention )

  (* PRESSURE monitoring block - indication, no set-point invented )
  FB_AI_QUAIL_CAGEPT-01( PV := QUAIL_CAGEPT-01_PV );
  QUAIL_CAGEPT-01_ALARM_HI := 9.0 ;  (* 90 % of span, registered LSH convention )

  (* TEMPERATURE monitoring block - indication, no set-point invented )
  FB_AI_QUAIL_CAGETE-01( PV := QUAIL_CAGETE-01_PV );
  QUAIL_CAGETE-01_ALARM_HI := 135.0 ;  (* 90 % of span, registered LSH convention )

  (* PRESSURE monitoring block - indication, no set-point invented )
  FB_AI_CHICKEN_COOPPT-01( PV := CHICKEN_COOPPT-01_PV );
  CHICKEN_COOPPT-01_ALARM_HI := 9.0 ;  (* 90 % of span, registered LSH convention )

  (* TEMPERATURE monitoring block - indication, no set-point invented )
  FB_AI_CHICKEN_COOPTE-01( PV := CHICKEN_COOPTE-01_PV );
  CHICKEN_COOPTE-01_ALARM_HI := 135.0 ;  (* 90 % of span, registered LSH convention )

  (* PRESSURE monitoring block - indication, no set-point invented )
  FB_AI_FEED_PREPPT-01( PV := FEED_PREPPT-01_PV );
  FEED_PREPPT-01_ALARM_HI := 9.0 ;  (* 90 % of span, registered LSH convention )

  (* TEMPERATURE monitoring block - indication, no set-point invented )
  FB_AI_FEED_PREPTE-01( PV := FEED_PREPTE-01_PV );
  FEED_PREPTE-01_ALARM_HI := 135.0 ;  (* 90 % of span, registered LSH convention )

  (* PRESSURE monitoring block - indication, no set-point invented )
  FB_AI_AQUA_TANKPT-01( PV := AQUA_TANKPT-01_PV );
  AQUA_TANKPT-01_ALARM_HI := 9.0 ;  (* 90 % of span, registered LSH convention )

  (* TEMPERATURE monitoring block - indication, no set-point invented )
  FB_AI_AQUA_TANKTE-01( PV := AQUA_TANKTE-01_PV );
  AQUA_TANKTE-01_ALARM_HI := 135.0 ;  (* 90 % of span, registered LSH convention )

  (* PRESSURE monitoring block - indication, no set-point invented )
  FB_AI_GROWBED_APT-01( PV := GROWBED_APT-01_PV );
  GROWBED_APT-01_ALARM_HI := 9.0 ;  (* 90 % of span, registered LSH convention )

  (* TEMPERATURE monitoring block - indication, no set-point invented )
  FB_AI_GROWBED_ATE-01( PV := GROWBED_ATE-01_PV );
  GROWBED_ATE-01_ALARM_HI := 135.0 ;  (* 90 % of span, registered LSH convention )

  (* PRESSURE monitoring block - indication, no set-point invented )
  FB_AI_GROWBED_BPT-01( PV := GROWBED_BPT-01_PV );
  GROWBED_BPT-01_ALARM_HI := 9.0 ;  (* 90 % of span, registered LSH convention )

  (* TEMPERATURE monitoring block - indication, no set-point invented )
  FB_AI_GROWBED_BTE-01( PV := GROWBED_BTE-01_PV );
  GROWBED_BTE-01_ALARM_HI := 135.0 ;  (* 90 % of span, registered LSH convention )

  (* PRESSURE monitoring block - indication, no set-point invented )
  FB_AI_BEE_HIVEPT-01( PV := BEE_HIVEPT-01_PV );
  BEE_HIVEPT-01_ALARM_HI := 9.0 ;  (* 90 % of span, registered LSH convention )

  (* TEMPERATURE monitoring block - indication, no set-point invented )
  FB_AI_BEE_HIVETE-01( PV := BEE_HIVETE-01_PV );
  BEE_HIVETE-01_ALARM_HI := 135.0 ;  (* 90 % of span, registered LSH convention )

  (* PRESSURE monitoring block - indication, no set-point invented )
  FB_AI_RABBIT_HUTCHPT-01( PV := RABBIT_HUTCHPT-01_PV );
  RABBIT_HUTCHPT-01_ALARM_HI := 9.0 ;  (* 90 % of span, registered LSH convention )

  (* TEMPERATURE monitoring block - indication, no set-point invented )
  FB_AI_RABBIT_HUTCHTE-01( PV := RABBIT_HUTCHTE-01_PV );
  RABBIT_HUTCHTE-01_ALARM_HI := 135.0 ;  (* 90 % of span, registered LSH convention )

  (* PRESSURE monitoring block - indication, no set-point invented )
  FB_AI_DUCK_PENPT-01( PV := DUCK_PENPT-01_PV );
  DUCK_PENPT-01_ALARM_HI := 9.0 ;  (* 90 % of span, registered LSH convention )

  (* TEMPERATURE monitoring block - indication, no set-point invented )
  FB_AI_DUCK_PENTE-01( PV := DUCK_PENTE-01_PV );
  DUCK_PENTE-01_ALARM_HI := 135.0 ;  (* 90 % of span, registered LSH convention )

  (* PRESSURE monitoring block - indication, no set-point invented )
  FB_AI_FOOD_STOREPT-01( PV := FOOD_STOREPT-01_PV );
  FOOD_STOREPT-01_ALARM_HI := 9.0 ;  (* 90 % of span, registered LSH convention )

  (* TEMPERATURE monitoring block - indication, no set-point invented )
  FB_AI_FOOD_STORETE-01( PV := FOOD_STORETE-01_PV );
  FOOD_STORETE-01_ALARM_HI := 135.0 ;  (* 90 % of span, registered LSH convention )

  (* PRESSURE monitoring block - indication, no set-point invented )
  FB_AI_AQUA_UVPT-01( PV := AQUA_UVPT-01_PV );
  AQUA_UVPT-01_ALARM_HI := 9.0 ;  (* 90 % of span, registered LSH convention )

  (* TEMPERATURE monitoring block - indication, no set-point invented )
  FB_AI_AQUA_UVTE-01( PV := AQUA_UVTE-01_PV );
  AQUA_UVTE-01_ALARM_HI := 135.0 ;  (* 90 % of span, registered LSH convention )

  (* PRESSURE monitoring block - indication, no set-point invented )
  FB_AI_VERMI_BINPT-01( PV := VERMI_BINPT-01_PV );
  VERMI_BINPT-01_ALARM_HI := 9.0 ;  (* 90 % of span, registered LSH convention )

  (* TEMPERATURE monitoring block - indication, no set-point invented )
  FB_AI_VERMI_BINTE-01( PV := VERMI_BINTE-01_PV );
  VERMI_BINTE-01_ALARM_HI := 135.0 ;  (* 90 % of span, registered LSH convention )

  (* LEVEL monitoring block - indication, no set-point invented )
  FB_AI_FOOD_STORELT-01( PV := FOOD_STORELT-01_PV );
  FOOD_STORELT-01_ALARM_HI := 90.0 ;  (* 90 % of span, registered LSH convention )

  (* CARBON-DIOXIDE monitoring block - indication, no set-point invented )
  FB_AI_HYDRO_GROWAE-01( PV := HYDRO_GROWAE-01_PV );
  HYDRO_GROWAE-01_ALARM_HI := 4500.0 ;  (* 90 % of span, registered LSH convention )

  (* PRESSURE monitoring block - indication, no set-point invented )
  FB_AI_FEED_PREPPSH-01( PV := FEED_PREPPSH-01_PV );
  FEED_PREPPSH-01_ALARM_HI := 225.0 ;  (* 90 % of span, registered LSH convention )

  (* FLOW monitoring block - indication, no set-point invented )
  FB_AI_AQUA_UVFIT-01( PV := AQUA_UVFIT-01_PV );
  AQUA_UVFIT-01_ALARM_HI := 90.0 ;  (* 90 % of span, registered LSH convention )

  (* UV monitoring block - indication, no set-point invented )
  FB_AI_AQUA_UVUVT-01( PV := AQUA_UVUVT-01_PV );
  AQUA_UVUVT-01_ALARM_HI := 4.5 ;  (* 90 % of span, registered LSH convention )

  (* LEVEL monitoring block - indication, no set-point invented )
  FB_AI_GROWBED_ALT-01( PV := GROWBED_ALT-01_PV );
  GROWBED_ALT-01_ALARM_HI := 270.0 ;  (* 90 % of span, registered LSH convention )

  (* LEVEL monitoring block - indication, no set-point invented )
  FB_AI_GROWBED_BLT-01( PV := GROWBED_BLT-01_PV );
  GROWBED_BLT-01_ALARM_HI := 270.0 ;  (* 90 % of span, registered LSH convention )

END_PROGRAM

(* ---- PLC-FOUNDRY.st ---- *)
(* AQS-CTL-004 X-CTL-04: control program source, generated by flow_graph/control/plc_programs.py *)
(* Basis: AQS-CTL-001 INSTRUMENT_INDEX.csv, AQS-CTL-002 control architecture, graph set-points. *)
(* PLC-FOUNDRY: CPU single; IO counts AI 87 AO 0 DI 19 DO 1 (modules per AQS-CTL-002, 16-channel, 20 % spare) *)
PROGRAM PLC_FOUNDRY_CTRL
VAR
  (* 100 ms cyclic task per AQS-CTL-002 *)
  AL_POTPT-01_PV : REAL ;  (* no design pressure on the graph )
  AL_POTTE-01_PV : REAL ;  (* band by service )
  CAST_LINELT-01_PV : REAL ;  (* A-M-182 liquid height )
  CAST_LINEPT-01_PV : REAL ;  (* no design pressure on the graph )
  CAST_LINETE-01_PV : REAL ;  (* band by service )
  CA_POTLT-01_PV : REAL ;  (* A-M-182 liquid height )
  CA_POTPT-01_PV : REAL ;  (* no design pressure on the graph )
  CA_POTTE-01_PV : REAL ;  (* band by service )
  COMB_HEATPT-01_PV : REAL ;  (* no design pressure on the graph )
  COMB_HEATTE-01_PV : REAL ;  (* band by service )
  CONT_CASTLT-01_PV : REAL ;  (* A-M-182 liquid height )
  CONT_CASTPT-01_PV : REAL ;  (* no design pressure on the graph )
  CONT_CASTTE-01_PV : REAL ;  (* band by service )
  CR_CELLPT-01_PV : REAL ;  (* no design pressure on the graph )
  CR_CELLTE-01_PV : REAL ;  (* band by service )
  DRAWPT-01_PV : REAL ;  (* no design pressure on the graph )
  DRAWTE-01_PV : REAL ;  (* band by service )
  EXTRUDEPT-01_PV : REAL ;  (* no design pressure on the graph )
  EXTRUDETE-01_PV : REAL ;  (* band by service )
  FLUX_PREPPT-01_PV : REAL ;  (* no design pressure on the graph )
  FLUX_PREPTE-01_PV : REAL ;  (* band by service )
  IND_MELTFT-01_PV : REAL ;  (* IND_MELT_TO_CAST normal 0.12 L/h )
  IND_MELTFT-02_PV : REAL ;  (* IND_TO_CONT normal 0.96 L/h )
  IND_MELTFT-03_PV : REAL ;  (* IND_TO_ATOM normal 0.00 L/h )
  IND_MELTFT-04_PV : REAL ;  (* IND_TO_INV normal 0.08 L/h )
  IND_MELTPT-01_PV : REAL ;  (* no design pressure on the graph )
  IND_MELTTE-01_PV : REAL ;  (* band by service )
  INV_CASTLT-01_PV : REAL ;  (* A-M-182 liquid height )
  INV_CASTPT-01_PV : REAL ;  (* no design pressure on the graph )
  INV_CASTTE-01_PV : REAL ;  (* band by service )
  METAL_STOREPT-01_PV : REAL ;  (* no design pressure on the graph )
  METAL_STORETE-01_PV : REAL ;  (* band by service )
  MG_POTLT-01_PV : REAL ;  (* A-M-182 liquid height )
  MG_POTPT-01_PV : REAL ;  (* no design pressure on the graph )
  MG_POTTE-01_PV : REAL ;  (* band by service )
  MO_CELLPT-01_PV : REAL ;  (* no design pressure on the graph )
  MO_CELLTE-01_PV : REAL ;  (* band by service )
  ROLLPT-01_PV : REAL ;  (* no design pressure on the graph )
  ROLLTE-01_PV : REAL ;  (* band by service )
  SHELL_BREAKLT-01_PV : REAL ;  (* A-M-182 liquid height )
  SHELL_BREAKPT-01_PV : REAL ;  (* no design pressure on the graph )
  SHELL_BREAKTE-01_PV : REAL ;  (* band by service )
  SHELL_BUILDPT-01_PV : REAL ;  (* no design pressure on the graph )
  SHELL_BUILDTE-01_PV : REAL ;  (* band by service )
  SHELL_BURNOUTFT-01_PV : REAL ;  (* WAX_RECLAIM_TO_PATTERN normal 0.07 L/h )
  SHELL_BURNOUTFT-02_PV : REAL ;  (* WAX_TO_OIL normal 0.00 L/h )
  SHELL_BURNOUTFT-03_PV : REAL ;  (* IA-BURNOUT-VENT normal 0.01 L/h )
  SHELL_BURNOUTPT-01_PV : REAL ;  (* no design pressure on the graph )
  SHELL_BURNOUTTE-01_PV : REAL ;  (* design T 900.0 C )
  SINTERPT-01_PV : REAL ;  (* no design pressure on the graph )
  SINTERTE-01_PV : REAL ;  (* design T 1300.0 C )
  STOCK_OUTPT-01_PV : REAL ;  (* no design pressure on the graph )
  STOCK_OUTTE-01_PV : REAL ;  (* band by service )
  TI_CELLFT-01_PV : REAL ;  (* TI_CELL_CL2_TO_CRU normal 0.00 L/h )
  TI_CELLFT-02_PV : REAL ;  (* IA-MGCL2-KROLL normal 0.08 L/h )
  TI_CELLFT-03_PV : REAL ;  (* IA-KROLL-CO normal 0.02 L/h )
  TI_CELLPT-01_PV : REAL ;  (* no design pressure on the graph )
  TI_CELLTE-01_PV : REAL ;  (* band by service )
  VAC_CASTPT-01_PV : REAL ;  (* no design pressure on the graph )
  VAC_CASTTE-01_PV : REAL ;  (* band by service )
  VAC_INDPT-01_PV : REAL ;  (* no design pressure on the graph )
  VAC_INDTE-01_PV : REAL ;  (* band by service )
  WAX_PATTERNLT-01_PV : REAL ;  (* A-M-182 liquid height )
  WAX_PATTERNPT-01_PV : REAL ;  (* no design pressure on the graph )
  WAX_PATTERNTE-01_PV : REAL ;  (* band by service )
  AL_POTIT-01_PV : REAL ;  (* cell current: design I_A 749.96 A )
  CA_POTIT-01_PV : REAL ;  (* cell current: design I_A 2.75 A )
  CR_CELLIT-01_PV : REAL ;  (* cell current: design I_A 18.95 A )
  MG_POTIT-01_PV : REAL ;  (* cell current: design I_A 54.89 A )
  MO_CELLIT-01_PV : REAL ;  (* cell current: design I_A 2.57 A )
  AL_POTAE-01_PV : REAL ;  (* anode-gas Cl2 offtake: IA-CL2-SHIP 39.42 kg/d; AL_POT_CL2 recycle standby )
  CA_POTAE-01_PV : REAL ;  (* anode-gas Cl2 offtake: IA-CA-CL2-SHIP 0.10 kg/d )
  CR_CELLAE-01_PV : REAL ;  (* carbochlorination loop Cl2 (design chemistry); IA-CR-VENT CO 0.20 kg/d )
  MG_POTAE-01_PV : REAL ;  (* anode-gas Cl2 to the Kroll chlorinator: IA-CL2-MG-TI 1.48 kg/d )
  MO_CELLAE-01_PV : REAL ;  (* anode gas (Cl2 or O2) to CRU: MO_CELL_ANODE_GAS_TO_CRU )
  TI_CELLLT-01_PV : REAL ;  (* TiCl4 receiver between chlorinator and retort (design chemistry, AQS-BAL-KROLL) )
  RF_HEATTE-01_PV : REAL ;  (* equal-duty backup of the IND_MELT crucible class (design backup_of) )
  RES_HEATTE-01_PV : REAL ;  (* design T_C 900 C (reheat, N+1 of SHELL_BURNOUT/SINTER) )
  FORGEZT-01_PV : REAL ;  (* ram stroke: design ram_mm 200 )
  FORGETE-01_PV : REAL ;  (* open-die press stock temperature (N+1 of ROLL); no design T on the graph )
  FLUX_PREPLT-01_PV : REAL ;  (* flux hopper: design hopper_L 20 L )
  SHELL_BUILDLT-01_PV : REAL ;  (* slurry tank: design slurry_L 40 L )
  E_HEATTE-01_PV : REAL ;  (* resistance element temperature watch on the N+1 melt trim duty (X-LOC-09 placeho )
  IND_MELTTE-90 : BOOL ;  (* SIF watch input, routed to the safety CPU pair (AQS-CTL-003) *)
  SHELL_BURNOUTTE-90 : BOOL ;  (* SIF watch input, routed to the safety CPU pair (AQS-CTL-003) *)
  RES_HEATTE-90 : BOOL ;  (* SIF watch input, routed to the safety CPU pair (AQS-CTL-003) *)
  SINTERTE-90 : BOOL ;  (* SIF watch input, routed to the safety CPU pair (AQS-CTL-003) *)
END_VAR

  (* PRESSURE monitoring block - indication, no set-point invented )
  FB_AI_AL_POTPT-01( PV := AL_POTPT-01_PV );
  AL_POTPT-01_ALARM_HI := 9.0 ;  (* 90 % of span, registered LSH convention )

  (* TEMPERATURE monitoring block - indication, no set-point invented )
  FB_AI_AL_POTTE-01( PV := AL_POTTE-01_PV );
  AL_POTTE-01_ALARM_HI := 135.0 ;  (* 90 % of span, registered LSH convention )

  (* LEVEL monitoring block - indication, no set-point invented )
  FB_AI_CAST_LINELT-01( PV := CAST_LINELT-01_PV );
  CAST_LINELT-01_ALARM_HI := 90.0 ;  (* 90 % of span, registered LSH convention )

  (* PRESSURE monitoring block - indication, no set-point invented )
  FB_AI_CAST_LINEPT-01( PV := CAST_LINEPT-01_PV );
  CAST_LINEPT-01_ALARM_HI := 9.0 ;  (* 90 % of span, registered LSH convention )

  (* TEMPERATURE monitoring block - indication, no set-point invented )
  FB_AI_CAST_LINETE-01( PV := CAST_LINETE-01_PV );
  CAST_LINETE-01_ALARM_HI := 135.0 ;  (* 90 % of span, registered LSH convention )

  (* LEVEL monitoring block - indication, no set-point invented )
  FB_AI_CA_POTLT-01( PV := CA_POTLT-01_PV );
  CA_POTLT-01_ALARM_HI := 90.0 ;  (* 90 % of span, registered LSH convention )

  (* PRESSURE monitoring block - indication, no set-point invented )
  FB_AI_CA_POTPT-01( PV := CA_POTPT-01_PV );
  CA_POTPT-01_ALARM_HI := 9.0 ;  (* 90 % of span, registered LSH convention )

  (* TEMPERATURE monitoring block - indication, no set-point invented )
  FB_AI_CA_POTTE-01( PV := CA_POTTE-01_PV );
  CA_POTTE-01_ALARM_HI := 135.0 ;  (* 90 % of span, registered LSH convention )

  (* PRESSURE monitoring block - indication, no set-point invented )
  FB_AI_COMB_HEATPT-01( PV := COMB_HEATPT-01_PV );
  COMB_HEATPT-01_ALARM_HI := 9.0 ;  (* 90 % of span, registered LSH convention )

  (* TEMPERATURE monitoring block - indication, no set-point invented )
  FB_AI_COMB_HEATTE-01( PV := COMB_HEATTE-01_PV );
  COMB_HEATTE-01_ALARM_HI := 135.0 ;  (* 90 % of span, registered LSH convention )

  (* LEVEL monitoring block - indication, no set-point invented )
  FB_AI_CONT_CASTLT-01( PV := CONT_CASTLT-01_PV );
  CONT_CASTLT-01_ALARM_HI := 90.0 ;  (* 90 % of span, registered LSH convention )

  (* PRESSURE monitoring block - indication, no set-point invented )
  FB_AI_CONT_CASTPT-01( PV := CONT_CASTPT-01_PV );
  CONT_CASTPT-01_ALARM_HI := 9.0 ;  (* 90 % of span, registered LSH convention )

  (* TEMPERATURE monitoring block - indication, no set-point invented )
  FB_AI_CONT_CASTTE-01( PV := CONT_CASTTE-01_PV );
  CONT_CASTTE-01_ALARM_HI := 135.0 ;  (* 90 % of span, registered LSH convention )

  (* PRESSURE monitoring block - indication, no set-point invented )
  FB_AI_CR_CELLPT-01( PV := CR_CELLPT-01_PV );
  CR_CELLPT-01_ALARM_HI := 9.0 ;  (* 90 % of span, registered LSH convention )

  (* TEMPERATURE monitoring block - indication, no set-point invented )
  FB_AI_CR_CELLTE-01( PV := CR_CELLTE-01_PV );
  CR_CELLTE-01_ALARM_HI := 135.0 ;  (* 90 % of span, registered LSH convention )

  (* PRESSURE monitoring block - indication, no set-point invented )
  FB_AI_DRAWPT-01( PV := DRAWPT-01_PV );
  DRAWPT-01_ALARM_HI := 9.0 ;  (* 90 % of span, registered LSH convention )

  (* TEMPERATURE monitoring block - indication, no set-point invented )
  FB_AI_DRAWTE-01( PV := DRAWTE-01_PV );
  DRAWTE-01_ALARM_HI := 135.0 ;  (* 90 % of span, registered LSH convention )

  (* PRESSURE monitoring block - indication, no set-point invented )
  FB_AI_EXTRUDEPT-01( PV := EXTRUDEPT-01_PV );
  EXTRUDEPT-01_ALARM_HI := 9.0 ;  (* 90 % of span, registered LSH convention )

  (* TEMPERATURE monitoring block - indication, no set-point invented )
  FB_AI_EXTRUDETE-01( PV := EXTRUDETE-01_PV );
  EXTRUDETE-01_ALARM_HI := 135.0 ;  (* 90 % of span, registered LSH convention )

  (* PRESSURE monitoring block - indication, no set-point invented )
  FB_AI_FLUX_PREPPT-01( PV := FLUX_PREPPT-01_PV );
  FLUX_PREPPT-01_ALARM_HI := 9.0 ;  (* 90 % of span, registered LSH convention )

  (* TEMPERATURE monitoring block - indication, no set-point invented )
  FB_AI_FLUX_PREPTE-01( PV := FLUX_PREPTE-01_PV );
  FLUX_PREPTE-01_ALARM_HI := 135.0 ;  (* 90 % of span, registered LSH convention )

  (* FLOW control loop - set-point from the graph basis *)
  IND_MELTFT-01_SP := 0.12 ;  (* graph basis: IND_MELT_TO_CAST normal 0.12 L/h )
  FB_PI_IND_MELTFT-01( PV := IND_MELTFT-01_PV, SP := IND_MELTFT-01_SP );  (* PI per AQS-CTL-002; GAIN/KI entered at commissioning from the step test (AQS-COM-001 sec. 3), anti-windup clamp per this FB *)
  IND_MELTFT-01_ALARM_HI := 0.132 ;  (* SP x 1.1 margin, A-M-188 margin class *)
  IND_MELTFT-01_ALARM_LO := 0.108 ;

  (* FLOW control loop - set-point from the graph basis *)
  IND_MELTFT-02_SP := 0.96 ;  (* graph basis: IND_TO_CONT normal 0.96 L/h )
  FB_PI_IND_MELTFT-02( PV := IND_MELTFT-02_PV, SP := IND_MELTFT-02_SP );  (* PI per AQS-CTL-002; GAIN/KI entered at commissioning from the step test (AQS-COM-001 sec. 3), anti-windup clamp per this FB *)
  IND_MELTFT-02_ALARM_HI := 1.056 ;  (* SP x 1.1 margin, A-M-188 margin class *)
  IND_MELTFT-02_ALARM_LO := 0.864 ;

  (* FLOW control loop - set-point from the graph basis *)
  IND_MELTFT-03_SP := 0.0 ;  (* graph basis: IND_TO_ATOM normal 0.00 L/h )
  FB_PI_IND_MELTFT-03( PV := IND_MELTFT-03_PV, SP := IND_MELTFT-03_SP );  (* PI per AQS-CTL-002; GAIN/KI entered at commissioning from the step test (AQS-COM-001 sec. 3), anti-windup clamp per this FB *)
  IND_MELTFT-03_ALARM_HI := 0.0 ;  (* expected-zero state: any positive PV alarms )

  (* FLOW control loop - set-point from the graph basis *)
  IND_MELTFT-04_SP := 0.08 ;  (* graph basis: IND_TO_INV normal 0.08 L/h )
  FB_PI_IND_MELTFT-04( PV := IND_MELTFT-04_PV, SP := IND_MELTFT-04_SP );  (* PI per AQS-CTL-002; GAIN/KI entered at commissioning from the step test (AQS-COM-001 sec. 3), anti-windup clamp per this FB *)
  IND_MELTFT-04_ALARM_HI := 0.08800000000000001 ;  (* SP x 1.1 margin, A-M-188 margin class *)
  IND_MELTFT-04_ALARM_LO := 0.07200000000000001 ;

  (* PRESSURE monitoring block - indication, no set-point invented )
  FB_AI_IND_MELTPT-01( PV := IND_MELTPT-01_PV );
  IND_MELTPT-01_ALARM_HI := 9.0 ;  (* 90 % of span, registered LSH convention )

  (* TEMPERATURE monitoring block - indication, no set-point invented )
  FB_AI_IND_MELTTE-01( PV := IND_MELTTE-01_PV );
  IND_MELTTE-01_ALARM_HI := 540.0 ;  (* 90 % of span, registered LSH convention )

  (* LEVEL monitoring block - indication, no set-point invented )
  FB_AI_INV_CASTLT-01( PV := INV_CASTLT-01_PV );
  INV_CASTLT-01_ALARM_HI := 90.0 ;  (* 90 % of span, registered LSH convention )

  (* PRESSURE monitoring block - indication, no set-point invented )
  FB_AI_INV_CASTPT-01( PV := INV_CASTPT-01_PV );
  INV_CASTPT-01_ALARM_HI := 9.0 ;  (* 90 % of span, registered LSH convention )

  (* TEMPERATURE monitoring block - indication, no set-point invented )
  FB_AI_INV_CASTTE-01( PV := INV_CASTTE-01_PV );
  INV_CASTTE-01_ALARM_HI := 135.0 ;  (* 90 % of span, registered LSH convention )

  (* PRESSURE monitoring block - indication, no set-point invented )
  FB_AI_METAL_STOREPT-01( PV := METAL_STOREPT-01_PV );
  METAL_STOREPT-01_ALARM_HI := 9.0 ;  (* 90 % of span, registered LSH convention )

  (* TEMPERATURE monitoring block - indication, no set-point invented )
  FB_AI_METAL_STORETE-01( PV := METAL_STORETE-01_PV );
  METAL_STORETE-01_ALARM_HI := 135.0 ;  (* 90 % of span, registered LSH convention )

  (* LEVEL monitoring block - indication, no set-point invented )
  FB_AI_MG_POTLT-01( PV := MG_POTLT-01_PV );
  MG_POTLT-01_ALARM_HI := 90.0 ;  (* 90 % of span, registered LSH convention )

  (* PRESSURE monitoring block - indication, no set-point invented )
  FB_AI_MG_POTPT-01( PV := MG_POTPT-01_PV );
  MG_POTPT-01_ALARM_HI := 9.0 ;  (* 90 % of span, registered LSH convention )

  (* TEMPERATURE monitoring block - indication, no set-point invented )
  FB_AI_MG_POTTE-01( PV := MG_POTTE-01_PV );
  MG_POTTE-01_ALARM_HI := 135.0 ;  (* 90 % of span, registered LSH convention )

  (* PRESSURE monitoring block - indication, no set-point invented )
  FB_AI_MO_CELLPT-01( PV := MO_CELLPT-01_PV );
  MO_CELLPT-01_ALARM_HI := 9.0 ;  (* 90 % of span, registered LSH convention )

  (* TEMPERATURE monitoring block - indication, no set-point invented )
  FB_AI_MO_CELLTE-01( PV := MO_CELLTE-01_PV );
  MO_CELLTE-01_ALARM_HI := 135.0 ;  (* 90 % of span, registered LSH convention )

  (* PRESSURE monitoring block - indication, no set-point invented )
  FB_AI_ROLLPT-01( PV := ROLLPT-01_PV );
  ROLLPT-01_ALARM_HI := 9.0 ;  (* 90 % of span, registered LSH convention )

  (* TEMPERATURE monitoring block - indication, no set-point invented )
  FB_AI_ROLLTE-01( PV := ROLLTE-01_PV );
  ROLLTE-01_ALARM_HI := 135.0 ;  (* 90 % of span, registered LSH convention )

  (* LEVEL monitoring block - indication, no set-point invented )
  FB_AI_SHELL_BREAKLT-01( PV := SHELL_BREAKLT-01_PV );
  SHELL_BREAKLT-01_ALARM_HI := 90.0 ;  (* 90 % of span, registered LSH convention )

  (* PRESSURE monitoring block - indication, no set-point invented )
  FB_AI_SHELL_BREAKPT-01( PV := SHELL_BREAKPT-01_PV );
  SHELL_BREAKPT-01_ALARM_HI := 9.0 ;  (* 90 % of span, registered LSH convention )

  (* TEMPERATURE monitoring block - indication, no set-point invented )
  FB_AI_SHELL_BREAKTE-01( PV := SHELL_BREAKTE-01_PV );
  SHELL_BREAKTE-01_ALARM_HI := 135.0 ;  (* 90 % of span, registered LSH convention )

  (* PRESSURE monitoring block - indication, no set-point invented )
  FB_AI_SHELL_BUILDPT-01( PV := SHELL_BUILDPT-01_PV );
  SHELL_BUILDPT-01_ALARM_HI := 9.0 ;  (* 90 % of span, registered LSH convention )

  (* TEMPERATURE monitoring block - indication, no set-point invented )
  FB_AI_SHELL_BUILDTE-01( PV := SHELL_BUILDTE-01_PV );
  SHELL_BUILDTE-01_ALARM_HI := 135.0 ;  (* 90 % of span, registered LSH convention )

  (* FLOW control loop - set-point from the graph basis *)
  SHELL_BURNOUTFT-01_SP := 0.07 ;  (* graph basis: WAX_RECLAIM_TO_PATTERN normal 0.07 L/h )
  FB_PI_SHELL_BURNOUTFT-01( PV := SHELL_BURNOUTFT-01_PV, SP := SHELL_BURNOUTFT-01_SP );  (* PI per AQS-CTL-002; GAIN/KI entered at commissioning from the step test (AQS-COM-001 sec. 3), anti-windup clamp per this FB *)
  SHELL_BURNOUTFT-01_ALARM_HI := 0.07700000000000001 ;  (* SP x 1.1 margin, A-M-188 margin class *)
  SHELL_BURNOUTFT-01_ALARM_LO := 0.06300000000000001 ;

  (* FLOW control loop - set-point from the graph basis *)
  SHELL_BURNOUTFT-02_SP := 0.0 ;  (* graph basis: WAX_TO_OIL normal 0.00 L/h )
  FB_PI_SHELL_BURNOUTFT-02( PV := SHELL_BURNOUTFT-02_PV, SP := SHELL_BURNOUTFT-02_SP );  (* PI per AQS-CTL-002; GAIN/KI entered at commissioning from the step test (AQS-COM-001 sec. 3), anti-windup clamp per this FB *)
  SHELL_BURNOUTFT-02_ALARM_HI := 0.0 ;  (* expected-zero state: any positive PV alarms )

  (* FLOW control loop - set-point from the graph basis *)
  SHELL_BURNOUTFT-03_SP := 0.01 ;  (* graph basis: IA-BURNOUT-VENT normal 0.01 L/h )
  FB_PI_SHELL_BURNOUTFT-03( PV := SHELL_BURNOUTFT-03_PV, SP := SHELL_BURNOUTFT-03_SP );  (* PI per AQS-CTL-002; GAIN/KI entered at commissioning from the step test (AQS-COM-001 sec. 3), anti-windup clamp per this FB *)
  SHELL_BURNOUTFT-03_ALARM_HI := 0.011000000000000001 ;  (* SP x 1.1 margin, A-M-188 margin class *)
  SHELL_BURNOUTFT-03_ALARM_LO := 0.009000000000000001 ;

  (* PRESSURE monitoring block - indication, no set-point invented )
  FB_AI_SHELL_BURNOUTPT-01( PV := SHELL_BURNOUTPT-01_PV );
  SHELL_BURNOUTPT-01_ALARM_HI := 9.0 ;  (* 90 % of span, registered LSH convention )

  (* TEMPERATURE control loop - set-point from the graph basis *)
  SHELL_BURNOUTTE-01_SP := 900.0 ;  (* graph basis: design T 900.0 C )
  FB_PI_SHELL_BURNOUTTE-01( PV := SHELL_BURNOUTTE-01_PV, SP := SHELL_BURNOUTTE-01_SP );  (* PI per AQS-CTL-002; GAIN/KI entered at commissioning from the step test (AQS-COM-001 sec. 3), anti-windup clamp per this FB *)
  SHELL_BURNOUTTE-01_ALARM_HI := 990.0000000000001 ;  (* SP x 1.1 margin, A-M-188 margin class *)
  SHELL_BURNOUTTE-01_ALARM_LO := 810.0 ;

  (* PRESSURE monitoring block - indication, no set-point invented )
  FB_AI_SINTERPT-01( PV := SINTERPT-01_PV );
  SINTERPT-01_ALARM_HI := 9.0 ;  (* 90 % of span, registered LSH convention )

  (* TEMPERATURE control loop - set-point from the graph basis *)
  SINTERTE-01_SP := 1300.0 ;  (* graph basis: design T 1300.0 C )
  FB_PI_SINTERTE-01( PV := SINTERTE-01_PV, SP := SINTERTE-01_SP );  (* PI per AQS-CTL-002; GAIN/KI entered at commissioning from the step test (AQS-COM-001 sec. 3), anti-windup clamp per this FB *)
  SINTERTE-01_ALARM_HI := 1430.0000000000002 ;  (* SP x 1.1 margin, A-M-188 margin class *)
  SINTERTE-01_ALARM_LO := 1170.0 ;

  (* PRESSURE monitoring block - indication, no set-point invented )
  FB_AI_STOCK_OUTPT-01( PV := STOCK_OUTPT-01_PV );
  STOCK_OUTPT-01_ALARM_HI := 9.0 ;  (* 90 % of span, registered LSH convention )

  (* TEMPERATURE monitoring block - indication, no set-point invented )
  FB_AI_STOCK_OUTTE-01( PV := STOCK_OUTTE-01_PV );
  STOCK_OUTTE-01_ALARM_HI := 135.0 ;  (* 90 % of span, registered LSH convention )

  (* FLOW control loop - set-point from the graph basis *)
  TI_CELLFT-01_SP := 0.0 ;  (* graph basis: TI_CELL_CL2_TO_CRU normal 0.00 L/h )
  FB_PI_TI_CELLFT-01( PV := TI_CELLFT-01_PV, SP := TI_CELLFT-01_SP );  (* PI per AQS-CTL-002; GAIN/KI entered at commissioning from the step test (AQS-COM-001 sec. 3), anti-windup clamp per this FB *)
  TI_CELLFT-01_ALARM_HI := 0.0 ;  (* expected-zero state: any positive PV alarms )

  (* FLOW control loop - set-point from the graph basis *)
  TI_CELLFT-02_SP := 0.08 ;  (* graph basis: IA-MGCL2-KROLL normal 0.08 L/h )
  FB_PI_TI_CELLFT-02( PV := TI_CELLFT-02_PV, SP := TI_CELLFT-02_SP );  (* PI per AQS-CTL-002; GAIN/KI entered at commissioning from the step test (AQS-COM-001 sec. 3), anti-windup clamp per this FB *)
  TI_CELLFT-02_ALARM_HI := 0.08800000000000001 ;  (* SP x 1.1 margin, A-M-188 margin class *)
  TI_CELLFT-02_ALARM_LO := 0.07200000000000001 ;

  (* FLOW control loop - set-point from the graph basis *)
  TI_CELLFT-03_SP := 0.02 ;  (* graph basis: IA-KROLL-CO normal 0.02 L/h )
  FB_PI_TI_CELLFT-03( PV := TI_CELLFT-03_PV, SP := TI_CELLFT-03_SP );  (* PI per AQS-CTL-002; GAIN/KI entered at commissioning from the step test (AQS-COM-001 sec. 3), anti-windup clamp per this FB *)
  TI_CELLFT-03_ALARM_HI := 0.022000000000000002 ;  (* SP x 1.1 margin, A-M-188 margin class *)
  TI_CELLFT-03_ALARM_LO := 0.018000000000000002 ;

  (* PRESSURE monitoring block - indication, no set-point invented )
  FB_AI_TI_CELLPT-01( PV := TI_CELLPT-01_PV );
  TI_CELLPT-01_ALARM_HI := 9.0 ;  (* 90 % of span, registered LSH convention )

  (* TEMPERATURE monitoring block - indication, no set-point invented )
  FB_AI_TI_CELLTE-01( PV := TI_CELLTE-01_PV );
  TI_CELLTE-01_ALARM_HI := 135.0 ;  (* 90 % of span, registered LSH convention )

  (* PRESSURE monitoring block - indication, no set-point invented )
  FB_AI_VAC_CASTPT-01( PV := VAC_CASTPT-01_PV );
  VAC_CASTPT-01_ALARM_HI := 9.0 ;  (* 90 % of span, registered LSH convention )

  (* TEMPERATURE monitoring block - indication, no set-point invented )
  FB_AI_VAC_CASTTE-01( PV := VAC_CASTTE-01_PV );
  VAC_CASTTE-01_ALARM_HI := 135.0 ;  (* 90 % of span, registered LSH convention )

  (* PRESSURE monitoring block - indication, no set-point invented )
  FB_AI_VAC_INDPT-01( PV := VAC_INDPT-01_PV );
  VAC_INDPT-01_ALARM_HI := 9.0 ;  (* 90 % of span, registered LSH convention )

  (* TEMPERATURE monitoring block - indication, no set-point invented )
  FB_AI_VAC_INDTE-01( PV := VAC_INDTE-01_PV );
  VAC_INDTE-01_ALARM_HI := 135.0 ;  (* 90 % of span, registered LSH convention )

  (* LEVEL monitoring block - indication, no set-point invented )
  FB_AI_WAX_PATTERNLT-01( PV := WAX_PATTERNLT-01_PV );
  WAX_PATTERNLT-01_ALARM_HI := 90.0 ;  (* 90 % of span, registered LSH convention )

  (* PRESSURE monitoring block - indication, no set-point invented )
  FB_AI_WAX_PATTERNPT-01( PV := WAX_PATTERNPT-01_PV );
  WAX_PATTERNPT-01_ALARM_HI := 9.0 ;  (* 90 % of span, registered LSH convention )

  (* TEMPERATURE monitoring block - indication, no set-point invented )
  FB_AI_WAX_PATTERNTE-01( PV := WAX_PATTERNTE-01_PV );
  WAX_PATTERNTE-01_ALARM_HI := 135.0 ;  (* 90 % of span, registered LSH convention )

  (* CURRENT control loop - set-point from the graph basis *)
  AL_POTIT-01_SP := 749.96 ;  (* graph basis: cell current: design I_A 749.96 A )
  FB_PI_AL_POTIT-01( PV := AL_POTIT-01_PV, SP := AL_POTIT-01_SP );  (* PI per AQS-CTL-002; GAIN/KI entered at commissioning from the step test (AQS-COM-001 sec. 3), anti-windup clamp per this FB *)
  AL_POTIT-01_ALARM_HI := 824.9560000000001 ;  (* SP x 1.1 margin, A-M-188 margin class *)
  AL_POTIT-01_ALARM_LO := 674.964 ;

  (* CURRENT control loop - set-point from the graph basis *)
  CA_POTIT-01_SP := 2.75 ;  (* graph basis: cell current: design I_A 2.75 A )
  FB_PI_CA_POTIT-01( PV := CA_POTIT-01_PV, SP := CA_POTIT-01_SP );  (* PI per AQS-CTL-002; GAIN/KI entered at commissioning from the step test (AQS-COM-001 sec. 3), anti-windup clamp per this FB *)
  CA_POTIT-01_ALARM_HI := 3.0250000000000004 ;  (* SP x 1.1 margin, A-M-188 margin class *)
  CA_POTIT-01_ALARM_LO := 2.475 ;

  (* CURRENT control loop - set-point from the graph basis *)
  CR_CELLIT-01_SP := 18.95 ;  (* graph basis: cell current: design I_A 18.95 A )
  FB_PI_CR_CELLIT-01( PV := CR_CELLIT-01_PV, SP := CR_CELLIT-01_SP );  (* PI per AQS-CTL-002; GAIN/KI entered at commissioning from the step test (AQS-COM-001 sec. 3), anti-windup clamp per this FB *)
  CR_CELLIT-01_ALARM_HI := 20.845000000000002 ;  (* SP x 1.1 margin, A-M-188 margin class *)
  CR_CELLIT-01_ALARM_LO := 17.055 ;

  (* CURRENT control loop - set-point from the graph basis *)
  MG_POTIT-01_SP := 54.89 ;  (* graph basis: cell current: design I_A 54.89 A )
  FB_PI_MG_POTIT-01( PV := MG_POTIT-01_PV, SP := MG_POTIT-01_SP );  (* PI per AQS-CTL-002; GAIN/KI entered at commissioning from the step test (AQS-COM-001 sec. 3), anti-windup clamp per this FB *)
  MG_POTIT-01_ALARM_HI := 60.379000000000005 ;  (* SP x 1.1 margin, A-M-188 margin class *)
  MG_POTIT-01_ALARM_LO := 49.401 ;

  (* CURRENT control loop - set-point from the graph basis *)
  MO_CELLIT-01_SP := 2.57 ;  (* graph basis: cell current: design I_A 2.57 A )
  FB_PI_MO_CELLIT-01( PV := MO_CELLIT-01_PV, SP := MO_CELLIT-01_SP );  (* PI per AQS-CTL-002; GAIN/KI entered at commissioning from the step test (AQS-COM-001 sec. 3), anti-windup clamp per this FB *)
  MO_CELLIT-01_ALARM_HI := 2.827 ;  (* SP x 1.1 margin, A-M-188 margin class *)
  MO_CELLIT-01_ALARM_LO := 2.3129999999999997 ;

  (* CHLORINE monitoring block - indication, no set-point invented )
  FB_AI_AL_POTAE-01( PV := AL_POTAE-01_PV );
  AL_POTAE-01_ALARM_HI := 90.0 ;  (* 90 % of span, registered LSH convention )

  (* CHLORINE monitoring block - indication, no set-point invented )
  FB_AI_CA_POTAE-01( PV := CA_POTAE-01_PV );
  CA_POTAE-01_ALARM_HI := 90.0 ;  (* 90 % of span, registered LSH convention )

  (* CHLORINE monitoring block - indication, no set-point invented )
  FB_AI_CR_CELLAE-01( PV := CR_CELLAE-01_PV );
  CR_CELLAE-01_ALARM_HI := 90.0 ;  (* 90 % of span, registered LSH convention )

  (* CHLORINE monitoring block - indication, no set-point invented )
  FB_AI_MG_POTAE-01( PV := MG_POTAE-01_PV );
  MG_POTAE-01_ALARM_HI := 90.0 ;  (* 90 % of span, registered LSH convention )

  (* CHLORINE monitoring block - indication, no set-point invented )
  FB_AI_MO_CELLAE-01( PV := MO_CELLAE-01_PV );
  MO_CELLAE-01_ALARM_HI := 90.0 ;  (* 90 % of span, registered LSH convention )

  (* LEVEL monitoring block - indication, no set-point invented )
  FB_AI_TI_CELLLT-01( PV := TI_CELLLT-01_PV );
  TI_CELLLT-01_ALARM_HI := 90.0 ;  (* 90 % of span, registered LSH convention )

  (* TEMPERATURE monitoring block - indication, no set-point invented )
  FB_AI_RF_HEATTE-01( PV := RF_HEATTE-01_PV );
  RF_HEATTE-01_ALARM_HI := 1440.0 ;  (* 90 % of span, registered LSH convention )

  (* TEMPERATURE control loop - set-point from the graph basis *)
  RES_HEATTE-01_SP := 900.0 ;  (* graph basis: design T_C 900 C (reheat, N+1 of SHELL_BURNOUT/SINTER) )
  FB_PI_RES_HEATTE-01( PV := RES_HEATTE-01_PV, SP := RES_HEATTE-01_SP );  (* PI per AQS-CTL-002; GAIN/KI entered at commissioning from the step test (AQS-COM-001 sec. 3), anti-windup clamp per this FB *)
  RES_HEATTE-01_ALARM_HI := 990.0000000000001 ;  (* SP x 1.1 margin, A-M-188 margin class *)
  RES_HEATTE-01_ALARM_LO := 810.0 ;

  (* POSITION monitoring block - indication, no set-point invented )
  FB_AI_FORGEZT-01( PV := FORGEZT-01_PV );
  FORGEZT-01_ALARM_HI := 180.0 ;  (* 90 % of span, registered LSH convention )

  (* TEMPERATURE monitoring block - indication, no set-point invented )
  FB_AI_FORGETE-01( PV := FORGETE-01_PV );
  FORGETE-01_ALARM_HI := 540.0 ;  (* 90 % of span, registered LSH convention )

  (* LEVEL monitoring block - indication, no set-point invented )
  FB_AI_FLUX_PREPLT-01( PV := FLUX_PREPLT-01_PV );
  FLUX_PREPLT-01_ALARM_HI := 90.0 ;  (* 90 % of span, registered LSH convention )

  (* LEVEL monitoring block - indication, no set-point invented )
  FB_AI_SHELL_BUILDLT-01( PV := SHELL_BUILDLT-01_PV );
  SHELL_BUILDLT-01_ALARM_HI := 90.0 ;  (* 90 % of span, registered LSH convention )

  (* TEMPERATURE monitoring block - indication, no set-point invented )
  FB_AI_E_HEATTE-01( PV := E_HEATTE-01_PV );
  E_HEATTE-01_ALARM_HI := 540.0 ;  (* 90 % of span, registered LSH convention )

  (* SIF watch passthrough, no action in the basic program )
  SIF_WATCH_IND_MELTTE-90 := IND_MELTTE-90 ;  (* to safety CPU pair, AQS-CTL-003 )

  (* SIF watch passthrough, no action in the basic program )
  SIF_WATCH_SHELL_BURNOUTTE-90 := SHELL_BURNOUTTE-90 ;  (* to safety CPU pair, AQS-CTL-003 )

  (* SIF watch passthrough, no action in the basic program )
  SIF_WATCH_RES_HEATTE-90 := RES_HEATTE-90 ;  (* to safety CPU pair, AQS-CTL-003 )

  (* SIF watch passthrough, no action in the basic program )
  SIF_WATCH_SINTERTE-90 := SINTERTE-90 ;  (* to safety CPU pair, AQS-CTL-003 )

END_PROGRAM

(* ---- PLC-GAS.st ---- *)
(* AQS-CTL-004 X-CTL-04: control program source, generated by flow_graph/control/plc_programs.py *)
(* Basis: AQS-CTL-001 INSTRUMENT_INDEX.csv, AQS-CTL-002 control architecture, graph set-points. *)
(* PLC-GAS: CPU redundant pair; IO counts AI 32 AO 0 DI 34 DO 6 (modules per AQS-CTL-002, 16-channel, 20 % spare) *)
PROGRAM PLC_GAS_CTRL
VAR
  (* 100 ms cyclic task per AQS-CTL-002 *)
  ACID_POLISH_SCRUBFT-01_PV : REAL ;  (* S66 normal 1.14 L/h )
  ACID_POLISH_SCRUBFT-02_PV : REAL ;  (* IA-ACID-AIR-RET normal 1562.91 L/h )
  ACID_POLISH_SCRUBLT-01_PV : REAL ;  (* A-M-182 liquid height )
  ACID_POLISH_SCRUBPT-01_PV : REAL ;  (* no design pressure on the graph )
  ACID_POLISH_SCRUBTE-01_PV : REAL ;  (* band by service )
  AFTERBURNER_FLUEPT-01_PV : REAL ;  (* no design pressure on the graph )
  AFTERBURNER_FLUETE-01_PV : REAL ;  (* band by service )
  ALK_SCRUBBERLT-01_PV : REAL ;  (* A-M-182 liquid height )
  ALK_SCRUBBERPT-01_PV : REAL ;  (* no design pressure on the graph )
  ALK_SCRUBBERTE-01_PV : REAL ;  (* band by service )
  BAGHOUSEFT-01_PV : REAL ;  (* IA-BAG-01 normal 0.30 L/h )
  BAGHOUSEPT-01_PV : REAL ;  (* no design pressure on the graph )
  BAGHOUSETE-01_PV : REAL ;  (* band by service )
  H2_DRYERLT-01_PV : REAL ;  (* A-M-182 liquid height )
  H2_DRYERPT-01_PV : REAL ;  (* no design pressure on the graph )
  H2_DRYERTE-01_PV : REAL ;  (* design T 250.0 C )
  NOX_SCRUBFT-01_PV : REAL ;  (* IA-NOX-H2O normal 9.22 L/h )
  NOX_SCRUBFT-02_PV : REAL ;  (* IA-NOX-N normal 0.84 L/h )
  NOX_SCRUBFT-03_PV : REAL ;  (* IA-NOX-CO2 normal 0.95 L/h )
  NOX_SCRUBFT-04_PV : REAL ;  (* IA-NOX-N2 normal 8.97 L/h )
  NOX_SCRUBLT-01_PV : REAL ;  (* A-M-182 liquid height )
  NOX_SCRUBPT-01_PV : REAL ;  (* no design pressure on the graph )
  NOX_SCRUBTE-01_PV : REAL ;  (* band by service )
  FLUE_KOLT-01_PV : REAL ;  (* A-M-182 liquid height )
  FLUE_KOPT-01_PV : REAL ;  (* no design pressure on the graph )
  FLUE_KOTE-01_PV : REAL ;  (* band by service )
  HDR_H2PT-01_PV : REAL ;  (* H2 pool header: IA-HDR-H2-02 1.98 kg/d max feed; no design pressure on the graph )
  HDR_O2PT-01_PV : REAL ;  (* O2 pool header: S83 33.2 kg/d product + returns; no design pressure on the graph )
  ATM_INTPT-01_PV : REAL ;  (* compressor discharge pressure watch against the process pressure (X-LOC-09 place )
  REC_HDRPT-01_PV : REAL ;  (* recovery header pressure watch; the header takes every relief and offgas dischar )
  AFTERBURNER_FLUETE-90 : BOOL ;  (* SIF watch input, routed to the safety CPU pair (AQS-CTL-003) *)
  H2_DRYERTE-90 : BOOL ;  (* SIF watch input, routed to the safety CPU pair (AQS-CTL-003) *)
END_VAR

  (* FLOW control loop - set-point from the graph basis *)
  ACID_POLISH_SCRUBFT-01_SP := 1.14 ;  (* graph basis: S66 normal 1.14 L/h )
  FB_PI_ACID_POLISH_SCRUBFT-01( PV := ACID_POLISH_SCRUBFT-01_PV, SP := ACID_POLISH_SCRUBFT-01_SP );  (* PI per AQS-CTL-002; GAIN/KI entered at commissioning from the step test (AQS-COM-001 sec. 3), anti-windup clamp per this FB *)
  ACID_POLISH_SCRUBFT-01_ALARM_HI := 1.254 ;  (* SP x 1.1 margin, A-M-188 margin class *)
  ACID_POLISH_SCRUBFT-01_ALARM_LO := 1.026 ;

  (* FLOW control loop - set-point from the graph basis *)
  ACID_POLISH_SCRUBFT-02_SP := 1562.91 ;  (* graph basis: IA-ACID-AIR-RET normal 1562.91 L/h )
  FB_PI_ACID_POLISH_SCRUBFT-02( PV := ACID_POLISH_SCRUBFT-02_PV, SP := ACID_POLISH_SCRUBFT-02_SP );  (* PI per AQS-CTL-002; GAIN/KI entered at commissioning from the step test (AQS-COM-001 sec. 3), anti-windup clamp per this FB *)
  ACID_POLISH_SCRUBFT-02_ALARM_HI := 1719.2010000000002 ;  (* SP x 1.1 margin, A-M-188 margin class *)
  ACID_POLISH_SCRUBFT-02_ALARM_LO := 1406.6190000000001 ;

  (* LEVEL monitoring block - indication, no set-point invented )
  FB_AI_ACID_POLISH_SCRUBLT-01( PV := ACID_POLISH_SCRUBLT-01_PV );
  ACID_POLISH_SCRUBLT-01_ALARM_HI := 90.0 ;  (* 90 % of span, registered LSH convention )

  (* PRESSURE monitoring block - indication, no set-point invented )
  FB_AI_ACID_POLISH_SCRUBPT-01( PV := ACID_POLISH_SCRUBPT-01_PV );
  ACID_POLISH_SCRUBPT-01_ALARM_HI := 9.0 ;  (* 90 % of span, registered LSH convention )

  (* TEMPERATURE monitoring block - indication, no set-point invented )
  FB_AI_ACID_POLISH_SCRUBTE-01( PV := ACID_POLISH_SCRUBTE-01_PV );
  ACID_POLISH_SCRUBTE-01_ALARM_HI := 135.0 ;  (* 90 % of span, registered LSH convention )

  (* PRESSURE monitoring block - indication, no set-point invented )
  FB_AI_AFTERBURNER_FLUEPT-01( PV := AFTERBURNER_FLUEPT-01_PV );
  AFTERBURNER_FLUEPT-01_ALARM_HI := 9.0 ;  (* 90 % of span, registered LSH convention )

  (* TEMPERATURE monitoring block - indication, no set-point invented )
  FB_AI_AFTERBURNER_FLUETE-01( PV := AFTERBURNER_FLUETE-01_PV );
  AFTERBURNER_FLUETE-01_ALARM_HI := 540.0 ;  (* 90 % of span, registered LSH convention )

  (* LEVEL monitoring block - indication, no set-point invented )
  FB_AI_ALK_SCRUBBERLT-01( PV := ALK_SCRUBBERLT-01_PV );
  ALK_SCRUBBERLT-01_ALARM_HI := 90.0 ;  (* 90 % of span, registered LSH convention )

  (* PRESSURE monitoring block - indication, no set-point invented )
  FB_AI_ALK_SCRUBBERPT-01( PV := ALK_SCRUBBERPT-01_PV );
  ALK_SCRUBBERPT-01_ALARM_HI := 9.0 ;  (* 90 % of span, registered LSH convention )

  (* TEMPERATURE monitoring block - indication, no set-point invented )
  FB_AI_ALK_SCRUBBERTE-01( PV := ALK_SCRUBBERTE-01_PV );
  ALK_SCRUBBERTE-01_ALARM_HI := 135.0 ;  (* 90 % of span, registered LSH convention )

  (* FLOW control loop - set-point from the graph basis *)
  BAGHOUSEFT-01_SP := 0.3 ;  (* graph basis: IA-BAG-01 normal 0.30 L/h )
  FB_PI_BAGHOUSEFT-01( PV := BAGHOUSEFT-01_PV, SP := BAGHOUSEFT-01_SP );  (* PI per AQS-CTL-002; GAIN/KI entered at commissioning from the step test (AQS-COM-001 sec. 3), anti-windup clamp per this FB *)
  BAGHOUSEFT-01_ALARM_HI := 0.33 ;  (* SP x 1.1 margin, A-M-188 margin class *)
  BAGHOUSEFT-01_ALARM_LO := 0.27 ;

  (* PRESSURE monitoring block - indication, no set-point invented )
  FB_AI_BAGHOUSEPT-01( PV := BAGHOUSEPT-01_PV );
  BAGHOUSEPT-01_ALARM_HI := 9.0 ;  (* 90 % of span, registered LSH convention )

  (* TEMPERATURE monitoring block - indication, no set-point invented )
  FB_AI_BAGHOUSETE-01( PV := BAGHOUSETE-01_PV );
  BAGHOUSETE-01_ALARM_HI := 135.0 ;  (* 90 % of span, registered LSH convention )

  (* LEVEL monitoring block - indication, no set-point invented )
  FB_AI_H2_DRYERLT-01( PV := H2_DRYERLT-01_PV );
  H2_DRYERLT-01_ALARM_HI := 90.0 ;  (* 90 % of span, registered LSH convention )

  (* PRESSURE monitoring block - indication, no set-point invented )
  FB_AI_H2_DRYERPT-01( PV := H2_DRYERPT-01_PV );
  H2_DRYERPT-01_ALARM_HI := 9.0 ;  (* 90 % of span, registered LSH convention )

  (* TEMPERATURE control loop - set-point from the graph basis *)
  H2_DRYERTE-01_SP := 250.0 ;  (* graph basis: design T 250.0 C )
  FB_PI_H2_DRYERTE-01( PV := H2_DRYERTE-01_PV, SP := H2_DRYERTE-01_SP );  (* PI per AQS-CTL-002; GAIN/KI entered at commissioning from the step test (AQS-COM-001 sec. 3), anti-windup clamp per this FB *)
  H2_DRYERTE-01_ALARM_HI := 275.0 ;  (* SP x 1.1 margin, A-M-188 margin class *)
  H2_DRYERTE-01_ALARM_LO := 225.0 ;

  (* FLOW control loop - set-point from the graph basis *)
  NOX_SCRUBFT-01_SP := 9.22 ;  (* graph basis: IA-NOX-H2O normal 9.22 L/h )
  FB_PI_NOX_SCRUBFT-01( PV := NOX_SCRUBFT-01_PV, SP := NOX_SCRUBFT-01_SP );  (* PI per AQS-CTL-002; GAIN/KI entered at commissioning from the step test (AQS-COM-001 sec. 3), anti-windup clamp per this FB *)
  NOX_SCRUBFT-01_ALARM_HI := 10.142000000000001 ;  (* SP x 1.1 margin, A-M-188 margin class *)
  NOX_SCRUBFT-01_ALARM_LO := 8.298 ;

  (* FLOW control loop - set-point from the graph basis *)
  NOX_SCRUBFT-02_SP := 0.84 ;  (* graph basis: IA-NOX-N normal 0.84 L/h )
  FB_PI_NOX_SCRUBFT-02( PV := NOX_SCRUBFT-02_PV, SP := NOX_SCRUBFT-02_SP );  (* PI per AQS-CTL-002; GAIN/KI entered at commissioning from the step test (AQS-COM-001 sec. 3), anti-windup clamp per this FB *)
  NOX_SCRUBFT-02_ALARM_HI := 0.924 ;  (* SP x 1.1 margin, A-M-188 margin class *)
  NOX_SCRUBFT-02_ALARM_LO := 0.756 ;

  (* FLOW control loop - set-point from the graph basis *)
  NOX_SCRUBFT-03_SP := 0.95 ;  (* graph basis: IA-NOX-CO2 normal 0.95 L/h )
  FB_PI_NOX_SCRUBFT-03( PV := NOX_SCRUBFT-03_PV, SP := NOX_SCRUBFT-03_SP );  (* PI per AQS-CTL-002; GAIN/KI entered at commissioning from the step test (AQS-COM-001 sec. 3), anti-windup clamp per this FB *)
  NOX_SCRUBFT-03_ALARM_HI := 1.045 ;  (* SP x 1.1 margin, A-M-188 margin class *)
  NOX_SCRUBFT-03_ALARM_LO := 0.855 ;

  (* FLOW control loop - set-point from the graph basis *)
  NOX_SCRUBFT-04_SP := 8.97 ;  (* graph basis: IA-NOX-N2 normal 8.97 L/h )
  FB_PI_NOX_SCRUBFT-04( PV := NOX_SCRUBFT-04_PV, SP := NOX_SCRUBFT-04_SP );  (* PI per AQS-CTL-002; GAIN/KI entered at commissioning from the step test (AQS-COM-001 sec. 3), anti-windup clamp per this FB *)
  NOX_SCRUBFT-04_ALARM_HI := 9.867 ;  (* SP x 1.1 margin, A-M-188 margin class *)
  NOX_SCRUBFT-04_ALARM_LO := 8.073 ;

  (* LEVEL monitoring block - indication, no set-point invented )
  FB_AI_NOX_SCRUBLT-01( PV := NOX_SCRUBLT-01_PV );
  NOX_SCRUBLT-01_ALARM_HI := 90.0 ;  (* 90 % of span, registered LSH convention )

  (* PRESSURE monitoring block - indication, no set-point invented )
  FB_AI_NOX_SCRUBPT-01( PV := NOX_SCRUBPT-01_PV );
  NOX_SCRUBPT-01_ALARM_HI := 9.0 ;  (* 90 % of span, registered LSH convention )

  (* TEMPERATURE monitoring block - indication, no set-point invented )
  FB_AI_NOX_SCRUBTE-01( PV := NOX_SCRUBTE-01_PV );
  NOX_SCRUBTE-01_ALARM_HI := 135.0 ;  (* 90 % of span, registered LSH convention )

  (* LEVEL monitoring block - indication, no set-point invented )
  FB_AI_FLUE_KOLT-01( PV := FLUE_KOLT-01_PV );
  FLUE_KOLT-01_ALARM_HI := 90.0 ;  (* 90 % of span, registered LSH convention )

  (* PRESSURE monitoring block - indication, no set-point invented )
  FB_AI_FLUE_KOPT-01( PV := FLUE_KOPT-01_PV );
  FLUE_KOPT-01_ALARM_HI := 9.0 ;  (* 90 % of span, registered LSH convention )

  (* TEMPERATURE monitoring block - indication, no set-point invented )
  FB_AI_FLUE_KOTE-01( PV := FLUE_KOTE-01_PV );
  FLUE_KOTE-01_ALARM_HI := 135.0 ;  (* 90 % of span, registered LSH convention )

  (* PRESSURE monitoring block - indication, no set-point invented )
  FB_AI_HDR_H2PT-01( PV := HDR_H2PT-01_PV );
  HDR_H2PT-01_ALARM_HI := 9.0 ;  (* 90 % of span, registered LSH convention )

  (* PRESSURE monitoring block - indication, no set-point invented )
  FB_AI_HDR_O2PT-01( PV := HDR_O2PT-01_PV );
  HDR_O2PT-01_ALARM_HI := 9.0 ;  (* 90 % of span, registered LSH convention )

  (* PRESSURE monitoring block - indication, no set-point invented )
  FB_AI_ATM_INTPT-01( PV := ATM_INTPT-01_PV );
  ATM_INTPT-01_ALARM_HI := 360.0 ;  (* 90 % of span, registered LSH convention )

  (* PRESSURE monitoring block - indication, no set-point invented )
  FB_AI_REC_HDRPT-01( PV := REC_HDRPT-01_PV );
  REC_HDRPT-01_ALARM_HI := 360.0 ;  (* 90 % of span, registered LSH convention )

  (* SIF watch passthrough, no action in the basic program )
  SIF_WATCH_AFTERBURNER_FLUETE-90 := AFTERBURNER_FLUETE-90 ;  (* to safety CPU pair, AQS-CTL-003 )

  (* SIF watch passthrough, no action in the basic program )
  SIF_WATCH_H2_DRYERTE-90 := H2_DRYERTE-90 ;  (* to safety CPU pair, AQS-CTL-003 )

END_PROGRAM

(* ---- PLC-GEO.st ---- *)
(* AQS-CTL-004 X-CTL-04: control program source, generated by flow_graph/control/plc_programs.py *)
(* Basis: AQS-CTL-001 INSTRUMENT_INDEX.csv, AQS-CTL-002 control architecture, graph set-points. *)
(* PLC-GEO: CPU redundant pair; IO counts AI 9 AO 0 DI 6 DO 3 (modules per AQS-CTL-002, 16-channel, 20 % spare) *)
PROGRAM PLC_GEO_CTRL
VAR
  (* 100 ms cyclic task per AQS-CTL-002 *)
  GEO_HP_CLOSED_LOOPPT-01_PV : REAL ;  (* no design pressure on the graph )
  GEO_HP_CLOSED_LOOPTE-01_PV : REAL ;  (* band by service )
  GEO_GHEXFT-01_PV : REAL ;  (* S43 normal 0.00 L/h )
  GEO_GHEXPT-01_PV : REAL ;  (* no design pressure on the graph )
  GEO_GHEXTE-01_PV : REAL ;  (* band by service )
  GEO_HPPT-01_PV : REAL ;  (* no design pressure on the graph )
  GEO_HPTE-01_PV : REAL ;  (* band by service )
  GEO_ORCPT-01_PV : REAL ;  (* no design pressure on the graph )
  GEO_ORCTE-01_PV : REAL ;  (* band by service )
END_VAR

  (* PRESSURE monitoring block - indication, no set-point invented )
  FB_AI_GEO_HP_CLOSED_LOOPPT-01( PV := GEO_HP_CLOSED_LOOPPT-01_PV );
  GEO_HP_CLOSED_LOOPPT-01_ALARM_HI := 9.0 ;  (* 90 % of span, registered LSH convention )

  (* TEMPERATURE monitoring block - indication, no set-point invented )
  FB_AI_GEO_HP_CLOSED_LOOPTE-01( PV := GEO_HP_CLOSED_LOOPTE-01_PV );
  GEO_HP_CLOSED_LOOPTE-01_ALARM_HI := 135.0 ;  (* 90 % of span, registered LSH convention )

  (* FLOW control loop - set-point from the graph basis *)
  GEO_GHEXFT-01_SP := 0.0 ;  (* graph basis: S43 normal 0.00 L/h )
  FB_PI_GEO_GHEXFT-01( PV := GEO_GHEXFT-01_PV, SP := GEO_GHEXFT-01_SP );  (* PI per AQS-CTL-002; GAIN/KI entered at commissioning from the step test (AQS-COM-001 sec. 3), anti-windup clamp per this FB *)
  GEO_GHEXFT-01_ALARM_HI := 0.0 ;  (* expected-zero state: any positive PV alarms )

  (* PRESSURE monitoring block - indication, no set-point invented )
  FB_AI_GEO_GHEXPT-01( PV := GEO_GHEXPT-01_PV );
  GEO_GHEXPT-01_ALARM_HI := 9.0 ;  (* 90 % of span, registered LSH convention )

  (* TEMPERATURE monitoring block - indication, no set-point invented )
  FB_AI_GEO_GHEXTE-01( PV := GEO_GHEXTE-01_PV );
  GEO_GHEXTE-01_ALARM_HI := 135.0 ;  (* 90 % of span, registered LSH convention )

  (* PRESSURE monitoring block - indication, no set-point invented )
  FB_AI_GEO_HPPT-01( PV := GEO_HPPT-01_PV );
  GEO_HPPT-01_ALARM_HI := 9.0 ;  (* 90 % of span, registered LSH convention )

  (* TEMPERATURE monitoring block - indication, no set-point invented )
  FB_AI_GEO_HPTE-01( PV := GEO_HPTE-01_PV );
  GEO_HPTE-01_ALARM_HI := 135.0 ;  (* 90 % of span, registered LSH convention )

  (* PRESSURE monitoring block - indication, no set-point invented )
  FB_AI_GEO_ORCPT-01( PV := GEO_ORCPT-01_PV );
  GEO_ORCPT-01_ALARM_HI := 9.0 ;  (* 90 % of span, registered LSH convention )

  (* TEMPERATURE monitoring block - indication, no set-point invented )
  FB_AI_GEO_ORCTE-01( PV := GEO_ORCTE-01_PV );
  GEO_ORCTE-01_ALARM_HI := 135.0 ;  (* 90 % of span, registered LSH convention )

END_PROGRAM

(* ---- PLC-GLASS.st ---- *)
(* AQS-CTL-004 X-CTL-04: control program source, generated by flow_graph/control/plc_programs.py *)
(* Basis: AQS-CTL-001 INSTRUMENT_INDEX.csv, AQS-CTL-002 control architecture, graph set-points. *)
(* PLC-GLASS: CPU single; IO counts AI 15 AO 0 DI 7 DO 0 (modules per AQS-CTL-002, 16-channel, 20 % spare) *)
PROGRAM PLC_GLASS_CTRL
VAR
  (* 100 ms cyclic task per AQS-CTL-002 *)
  GLASS_DIGESTFT-01_PV : REAL ;  (* IA-DIG-LIQ normal 0.92 L/h )
  GLASS_DIGESTFT-02_PV : REAL ;  (* IA-SIL-SRC normal 0.14 L/h )
  GLASS_DIGESTLT-01_PV : REAL ;  (* A-M-182 liquid height )
  GLASS_DIGESTPT-01_PV : REAL ;  (* no design pressure on the graph )
  GLASS_DIGESTTE-01_PV : REAL ;  (* design T 85 C )
  SI_REDUCEPT-01_PV : REAL ;  (* no design pressure on the graph )
  SI_REDUCETE-01_PV : REAL ;  (* band by service )
  GLASS_BURNOUTPT-01_PV : REAL ;  (* no design pressure on the graph )
  GLASS_BURNOUTTE-01_PV : REAL ;  (* band by service )
  GLASS_MILLPT-01_PV : REAL ;  (* no design pressure on the graph )
  GLASS_MILLTE-01_PV : REAL ;  (* band by service )
  GLASS_RINSEPT-01_PV : REAL ;  (* no design pressure on the graph )
  GLASS_RINSETE-01_PV : REAL ;  (* band by service )
  SI_REFINEPT-01_PV : REAL ;  (* no design pressure on the graph )
  SI_REFINETE-01_PV : REAL ;  (* band by service )
END_VAR

  (* FLOW control loop - set-point from the graph basis *)
  GLASS_DIGESTFT-01_SP := 0.92 ;  (* graph basis: IA-DIG-LIQ normal 0.92 L/h )
  FB_PI_GLASS_DIGESTFT-01( PV := GLASS_DIGESTFT-01_PV, SP := GLASS_DIGESTFT-01_SP );  (* PI per AQS-CTL-002; GAIN/KI entered at commissioning from the step test (AQS-COM-001 sec. 3), anti-windup clamp per this FB *)
  GLASS_DIGESTFT-01_ALARM_HI := 1.0120000000000002 ;  (* SP x 1.1 margin, A-M-188 margin class *)
  GLASS_DIGESTFT-01_ALARM_LO := 0.8280000000000001 ;

  (* FLOW control loop - set-point from the graph basis *)
  GLASS_DIGESTFT-02_SP := 0.14 ;  (* graph basis: IA-SIL-SRC normal 0.14 L/h )
  FB_PI_GLASS_DIGESTFT-02( PV := GLASS_DIGESTFT-02_PV, SP := GLASS_DIGESTFT-02_SP );  (* PI per AQS-CTL-002; GAIN/KI entered at commissioning from the step test (AQS-COM-001 sec. 3), anti-windup clamp per this FB *)
  GLASS_DIGESTFT-02_ALARM_HI := 0.15400000000000003 ;  (* SP x 1.1 margin, A-M-188 margin class *)
  GLASS_DIGESTFT-02_ALARM_LO := 0.12600000000000003 ;

  (* LEVEL monitoring block - indication, no set-point invented )
  FB_AI_GLASS_DIGESTLT-01( PV := GLASS_DIGESTLT-01_PV );
  GLASS_DIGESTLT-01_ALARM_HI := 90.0 ;  (* 90 % of span, registered LSH convention )

  (* PRESSURE monitoring block - indication, no set-point invented )
  FB_AI_GLASS_DIGESTPT-01( PV := GLASS_DIGESTPT-01_PV );
  GLASS_DIGESTPT-01_ALARM_HI := 9.0 ;  (* 90 % of span, registered LSH convention )

  (* TEMPERATURE control loop - set-point from the graph basis *)
  GLASS_DIGESTTE-01_SP := 85.0 ;  (* graph basis: design T 85 C )
  FB_PI_GLASS_DIGESTTE-01( PV := GLASS_DIGESTTE-01_PV, SP := GLASS_DIGESTTE-01_SP );  (* PI per AQS-CTL-002; GAIN/KI entered at commissioning from the step test (AQS-COM-001 sec. 3), anti-windup clamp per this FB *)
  GLASS_DIGESTTE-01_ALARM_HI := 93.50000000000001 ;  (* SP x 1.1 margin, A-M-188 margin class *)
  GLASS_DIGESTTE-01_ALARM_LO := 76.5 ;

  (* PRESSURE monitoring block - indication, no set-point invented )
  FB_AI_SI_REDUCEPT-01( PV := SI_REDUCEPT-01_PV );
  SI_REDUCEPT-01_ALARM_HI := 9.0 ;  (* 90 % of span, registered LSH convention )

  (* TEMPERATURE monitoring block - indication, no set-point invented )
  FB_AI_SI_REDUCETE-01( PV := SI_REDUCETE-01_PV );
  SI_REDUCETE-01_ALARM_HI := 135.0 ;  (* 90 % of span, registered LSH convention )

  (* PRESSURE monitoring block - indication, no set-point invented )
  FB_AI_GLASS_BURNOUTPT-01( PV := GLASS_BURNOUTPT-01_PV );
  GLASS_BURNOUTPT-01_ALARM_HI := 9.0 ;  (* 90 % of span, registered LSH convention )

  (* TEMPERATURE monitoring block - indication, no set-point invented )
  FB_AI_GLASS_BURNOUTTE-01( PV := GLASS_BURNOUTTE-01_PV );
  GLASS_BURNOUTTE-01_ALARM_HI := 135.0 ;  (* 90 % of span, registered LSH convention )

  (* PRESSURE monitoring block - indication, no set-point invented )
  FB_AI_GLASS_MILLPT-01( PV := GLASS_MILLPT-01_PV );
  GLASS_MILLPT-01_ALARM_HI := 9.0 ;  (* 90 % of span, registered LSH convention )

  (* TEMPERATURE monitoring block - indication, no set-point invented )
  FB_AI_GLASS_MILLTE-01( PV := GLASS_MILLTE-01_PV );
  GLASS_MILLTE-01_ALARM_HI := 135.0 ;  (* 90 % of span, registered LSH convention )

  (* PRESSURE monitoring block - indication, no set-point invented )
  FB_AI_GLASS_RINSEPT-01( PV := GLASS_RINSEPT-01_PV );
  GLASS_RINSEPT-01_ALARM_HI := 9.0 ;  (* 90 % of span, registered LSH convention )

  (* TEMPERATURE monitoring block - indication, no set-point invented )
  FB_AI_GLASS_RINSETE-01( PV := GLASS_RINSETE-01_PV );
  GLASS_RINSETE-01_ALARM_HI := 135.0 ;  (* 90 % of span, registered LSH convention )

  (* PRESSURE monitoring block - indication, no set-point invented )
  FB_AI_SI_REFINEPT-01( PV := SI_REFINEPT-01_PV );
  SI_REFINEPT-01_ALARM_HI := 9.0 ;  (* 90 % of span, registered LSH convention )

  (* TEMPERATURE monitoring block - indication, no set-point invented )
  FB_AI_SI_REFINETE-01( PV := SI_REFINETE-01_PV );
  SI_REFINETE-01_ALARM_HI := 135.0 ;  (* 90 % of span, registered LSH convention )

END_PROGRAM

(* ---- PLC-HAB.st ---- *)
(* AQS-CTL-004 X-CTL-04: control program source, generated by flow_graph/control/plc_programs.py *)
(* Basis: AQS-CTL-001 INSTRUMENT_INDEX.csv, AQS-CTL-002 control architecture, graph set-points. *)
(* PLC-HAB: CPU redundant pair; IO counts AI 13 AO 0 DI 1 DO 0 (modules per AQS-CTL-002, 16-channel, 20 % spare) *)
PROGRAM PLC_HAB_CTRL
VAR
  (* 100 ms cyclic task per AQS-CTL-002 *)
  HABITATIONLT-01_PV : REAL ;  (* A-M-182 liquid height )
  HABITATIONPT-01_PV : REAL ;  (* no design pressure on the graph )
  HABITATIONTE-01_PV : REAL ;  (* band by service )
  GALLEYPT-01_PV : REAL ;  (* no design pressure on the graph )
  GALLEYTE-01_PV : REAL ;  (* band by service )
  WASHROOMPT-01_PV : REAL ;  (* no design pressure on the graph )
  WASHROOMTE-01_PV : REAL ;  (* band by service )
  HDR_CO2PT-01_PV : REAL ;  (* CO2 header: S89 0.88 + S90 4.02 kg/d; no design pressure on the graph )
  HDR_N2PT-01_PV : REAL ;  (* plant air/N2 header: IA-AIR-RX-OUT 192.0 kg/d; no design pressure on the graph )
  COMMON_AREATE-01_PV : REAL ;  (* common-area temperature watch (X-HAB build-out; A-M-419) )
  MEDICALTE-01_PV : REAL ;  (* medical room temperature watch (X-HAB build-out; A-M-419) )
  REC_DAYROOMTE-01_PV : REAL ;  (* day-space temperature watch (X-HAB build-out; A-M-419) )
  SLEEP_QUARTERSTE-01_PV : REAL ;  (* quarters temperature watch (X-HAB build-out; A-M-419) )
END_VAR

  (* LEVEL monitoring block - indication, no set-point invented )
  FB_AI_HABITATIONLT-01( PV := HABITATIONLT-01_PV );
  HABITATIONLT-01_ALARM_HI := 90.0 ;  (* 90 % of span, registered LSH convention )

  (* PRESSURE monitoring block - indication, no set-point invented )
  FB_AI_HABITATIONPT-01( PV := HABITATIONPT-01_PV );
  HABITATIONPT-01_ALARM_HI := 9.0 ;  (* 90 % of span, registered LSH convention )

  (* TEMPERATURE monitoring block - indication, no set-point invented )
  FB_AI_HABITATIONTE-01( PV := HABITATIONTE-01_PV );
  HABITATIONTE-01_ALARM_HI := 135.0 ;  (* 90 % of span, registered LSH convention )

  (* PRESSURE monitoring block - indication, no set-point invented )
  FB_AI_GALLEYPT-01( PV := GALLEYPT-01_PV );
  GALLEYPT-01_ALARM_HI := 9.0 ;  (* 90 % of span, registered LSH convention )

  (* TEMPERATURE monitoring block - indication, no set-point invented )
  FB_AI_GALLEYTE-01( PV := GALLEYTE-01_PV );
  GALLEYTE-01_ALARM_HI := 135.0 ;  (* 90 % of span, registered LSH convention )

  (* PRESSURE monitoring block - indication, no set-point invented )
  FB_AI_WASHROOMPT-01( PV := WASHROOMPT-01_PV );
  WASHROOMPT-01_ALARM_HI := 9.0 ;  (* 90 % of span, registered LSH convention )

  (* TEMPERATURE monitoring block - indication, no set-point invented )
  FB_AI_WASHROOMTE-01( PV := WASHROOMTE-01_PV );
  WASHROOMTE-01_ALARM_HI := 135.0 ;  (* 90 % of span, registered LSH convention )

  (* PRESSURE monitoring block - indication, no set-point invented )
  FB_AI_HDR_CO2PT-01( PV := HDR_CO2PT-01_PV );
  HDR_CO2PT-01_ALARM_HI := 9.0 ;  (* 90 % of span, registered LSH convention )

  (* PRESSURE monitoring block - indication, no set-point invented )
  FB_AI_HDR_N2PT-01( PV := HDR_N2PT-01_PV );
  HDR_N2PT-01_ALARM_HI := 9.0 ;  (* 90 % of span, registered LSH convention )

  (* TEMPERATURE monitoring block - indication, no set-point invented )
  FB_AI_COMMON_AREATE-01( PV := COMMON_AREATE-01_PV );
  COMMON_AREATE-01_ALARM_HI := 135.0 ;  (* 90 % of span, registered LSH convention )

  (* TEMPERATURE monitoring block - indication, no set-point invented )
  FB_AI_MEDICALTE-01( PV := MEDICALTE-01_PV );
  MEDICALTE-01_ALARM_HI := 135.0 ;  (* 90 % of span, registered LSH convention )

  (* TEMPERATURE monitoring block - indication, no set-point invented )
  FB_AI_REC_DAYROOMTE-01( PV := REC_DAYROOMTE-01_PV );
  REC_DAYROOMTE-01_ALARM_HI := 135.0 ;  (* 90 % of span, registered LSH convention )

  (* TEMPERATURE monitoring block - indication, no set-point invented )
  FB_AI_SLEEP_QUARTERSTE-01( PV := SLEEP_QUARTERSTE-01_PV );
  SLEEP_QUARTERSTE-01_ALARM_HI := 135.0 ;  (* 90 % of span, registered LSH convention )

END_PROGRAM
